(* CODESYS project Example12_PLC.project

Project tree, tasks and I/O mapping:
  Device : CODESYS Control Win V3, 3S - Smart Software Solutions GmbH, order no. 305021, version 3.5.7.0
    application Application
      libraries: Standard, * (System)
      task MainTask (cyclic, interval t#20ms, priority 1) calls PLC_PRG
      program PLC_PRG [ST]
      global variables GVL
      function block FB_G4LTL [ST]
    Ethernet : Ethernet, 3S - Smart Software Solutions GmbH, version 3.5.7.0
      Modbus_TCP_Master : Modbus TCP Master, 3S - Smart Software Solutions GmbH, version 3.5.6.0
          settings: AutoReconnect = TRUE
        Modbus_TCP_Slave : Modbus TCP Slave, 3S - Smart Software Solutions GmbH, version 3.5.7.0
            settings: Unit-ID = 1; IPAddress = [127, 0, 0, 1]; Channel 0.Function Code = 4; Channel 0.Read Offset = 16#0000; Channel 0.Read Length = 1; Channel 0.Write Offset = 0; Channel 0.Write Length = 0; Channel 0.Cycle Time = 100; Channel 1.Function Code = 4; Channel 1.Read Offset = 16#0001; Channel 1.Read Length = 1; Channel 1.Write Offset = 0; Channel 1.Write Length = 0; Channel 1.Cycle Time = 100; Channel 2.Function Code = 4; Channel 2.Read Offset = 16#0002; Channel 2.Read Length = 1; Channel 2.Write Offset = 0; Channel 2.Write Length = 0; Channel 2.Cycle Time = 100; Channel 3.Function Code = 4; Channel 3.Read Offset = 16#0003; Channel 3.Read Length = 1; Channel 3.Write Offset = 0; Channel 3.Write Length = 0; Channel 3.Cycle Time = 100; Channel 4.Function Code = 4; Channel 4.Read Offset = 16#0004; Channel 4.Read Length = 1; Channel 4.Write Offset = 0; Channel 4.Write Length = 0; Channel 4.Cycle Time = 100; Channel 5.Function Code = 6; Channel 5.Read Offset = 0; Channel 5.Read Length = 0; Channel 5.Write Offset = 16#0000; Channel 5.Write Length = 1; Channel 5.Cycle Time = 100; Channel 6.Function Code = 6; Channel 6.Read Offset = 0;
              Channel 6.Read Length = 0; Channel 6.Write Offset = 16#0002; Channel 6.Write Length = 1; Channel 6.Cycle Time = 100; Channel 7.Function Code = 6; Channel 7.Read Offset = 0; Channel 7.Read Length = 0; Channel 7.Write Offset = 16#0003; Channel 7.Write Length = 1; Channel 7.Cycle Time = 100; Channel 8.Function Code = 6; Channel 8.Read Offset = 0; Channel 8.Read Length = 0; Channel 8.Write Offset = 16#0004; Channel 8.Write Length = 1; Channel 8.Cycle Time = 100; Channel 9.Function Code = 6; Channel 9.Read Offset = 0; Channel 9.Read Length = 0; Channel 9.Write Offset = 16#0001; Channel 9.Write Length = 1; Channel 9.Cycle Time = 100; Channel 10.Function Code = 4; Channel 10.Read Offset = 16#0005; Channel 10.Read Length = 1; Channel 10.Write Offset = 0; Channel 10.Write Length = 0; Channel 10.Cycle Time = 100
            input  Application.dIn0 : BOOL  // Channel 0.Channel 0.Bit0
            input  Application.dIn1 : BOOL  // Channel 1.Channel 1.Bit0
            input  Application.dIn2 : BOOL  // Channel 2.Channel 2.Bit0
            input  Application.dIn3 : BOOL  // Channel 3.Channel 3.Bit0
            input  Application.dIn4 : BOOL  // Channel 4.Channel 4.Bit0
            output Application.dOut0 : BOOL  // Channel 5.Channel 5.Bit0
            output Application.dOut2 : BOOL  // Channel 6.Channel 6.Bit0
            output Application.dOut3 : BOOL  // Channel 7.Channel 7.Bit0
            output Application.dOut4 : BOOL  // Channel 8.Channel 8.Bit0
            output Application.dOut1 : BOOL  // Channel 9.Channel 9.Bit0
            input  Application.dIn5 : BOOL  // Channel 10.Channel 10.Bit0
            unmapped channels: Channel 0, Channel 1, Channel 2, Channel 3, Channel 4, Channel 5, Channel 6, Channel 7, Channel 8, Channel 9, Channel 10
*)

// Device/Application/GVL
VAR_GLOBAL
	
dIn0 : BOOL;
dIn1 : BOOL;
dIn2 : BOOL;
dIn3 : BOOL;
dIn4 : BOOL;
dIn5 : BOOL;

dOut0 : BOOL;
dOut1 : BOOL; 
dOut2 : BOOL; 
dOut3 : BOOL; 
dOut4 : BOOL; 
END_VAR

// Device/Application/PLC_PRG
PROGRAM PLC_PRG
 

VAR 
	fb: FB_G4LTL;

	
END_VAR



// Direct looping
// Assign pins (from global variable to function block) 
fb.x0 := dIn0;
fb.x1 := dIn1;
fb.x2 := dIn2;
fb.x3 := dIn3;
fb.x4 := dIn4;
fb.x5 := dIn5;

// Assign pins (from function block to global variable)
dOut0 := fb.y0;
dOut1 := fb.y1;
dOut2 := fb.y2;

// Run the function block
fb();

END_PROGRAM

// Device/Application/FB_G4LTL
FUNCTION_BLOCK FB_G4LTL
   (* Variable definition *)
   VAR_INPUT
      x0	: BOOL;
      x1	: BOOL;
      x2	: BOOL;
      x3	: BOOL;
      x4	: BOOL;
      x5	: BOOL;
   END_VAR
   VAR_OUTPUT
      y0	: BOOL;
      y1	: BOOL;
      y2	: BOOL;
   END_VAR
   VAR
   (* The total number of states equals to 84 *)
      cstate98	: LINT := 0;
   END_VAR
   (* Constant definition  *)

 
   (* Control logic *)
CASE cstate98 OF
2090:
    IF ((x0 = FALSE) AND  (x1 = FALSE) AND  (x2 = FALSE) AND  (x3 = FALSE) AND  ( TRUE ) AND  (x5 = FALSE)) OR ((x0 = FALSE) AND  (x1 = FALSE) AND  (x2 = FALSE) AND  (x3 = TRUE) AND  (x4 = FALSE) AND  (x5 = FALSE)) THEN 
        cstate98 := 2122; y0 := FALSE; y1 := FALSE; y2 := FALSE;  
    ELSIF ((x0 = FALSE) AND  (x1 = FALSE) AND  (x2 = FALSE) AND  (x3 = FALSE) AND  ( TRUE ) AND  (x5 = TRUE)) OR ((x0 = FALSE) AND  (x1 = FALSE) AND  (x2 = FALSE) AND  (x3 = TRUE) AND  (x4 = FALSE) AND  (x5 = TRUE)) THEN 
        cstate98 := 2123; y0 := FALSE; y1 := FALSE; y2 := FALSE;  
    ELSIF ((x0 = FALSE) AND  (x1 = FALSE) AND  (x2 = FALSE) AND  (x3 = TRUE) AND  (x4 = TRUE) AND  ( TRUE )) THEN 
        cstate98 := 2090; y0 := FALSE; y1 := FALSE; y2 := FALSE;  
    ELSIF ((x0 = FALSE) AND  (x1 = FALSE) AND  (x2 = TRUE) AND  (x3 = FALSE) AND  ( TRUE ) AND  (x5 = FALSE)) THEN 
        cstate98 := 2602; y0 := FALSE; y1 := TRUE; y2 := FALSE;  
    ELSIF ((x0 = FALSE) AND  (x1 = FALSE) AND  (x2 = TRUE) AND  (x3 = FALSE) AND  ( TRUE ) AND  (x5 = TRUE)) THEN 
        cstate98 := 1610; y0 := FALSE; y1 := FALSE; y2 := FALSE;  
    ELSIF ((x0 = FALSE) AND  (x1 = FALSE) AND  (x2 = TRUE) AND  (x3 = TRUE) AND  ( TRUE ) AND  ( TRUE )) OR ((x0 = FALSE) AND  (x1 = TRUE) AND  (x2 = FALSE) AND  (x3 = TRUE) AND  ( TRUE ) AND  ( TRUE )) OR ((x0 = FALSE) AND  (x1 = TRUE) AND  (x2 = TRUE) AND  ( TRUE ) AND  ( TRUE ) AND  ( TRUE )) OR ((x0 = TRUE) AND  ( TRUE ) AND  (x2 = FALSE) AND  (x3 = TRUE) AND  ( TRUE ) AND  ( TRUE )) OR ((x0 = TRUE) AND  ( TRUE ) AND  (x2 = TRUE) AND  ( TRUE ) AND  ( TRUE ) AND  ( TRUE )) THEN 
        cstate98 := 617; y0 := FALSE; y1 := FALSE; y2 := FALSE;  
    ELSIF ((x0 = FALSE) AND  (x1 = TRUE) AND  (x2 = FALSE) AND  (x3 = FALSE) AND  ( TRUE ) AND  (x5 = FALSE)) OR ((x0 = TRUE) AND  ( TRUE ) AND  (x2 = FALSE) AND  (x3 = FALSE) AND  ( TRUE ) AND  (x5 = FALSE)) THEN 
        cstate98 := 3210; y0 := TRUE; y1 := FALSE; y2 := FALSE;  
    ELSIF ((x0 = FALSE) AND  (x1 = TRUE) AND  (x2 = FALSE) AND  (x3 = FALSE) AND  ( TRUE ) AND  (x5 = TRUE)) OR ((x0 = TRUE) AND  ( TRUE ) AND  (x2 = FALSE) AND  (x3 = FALSE) AND  ( TRUE ) AND  (x5 = TRUE)) THEN 
        cstate98 := 1194; y0 := FALSE; y1 := FALSE; y2 := FALSE;  
    END_IF;
2608:
    IF ((x0 = FALSE) AND  (x1 = FALSE) AND  (x2 = FALSE) AND  (x3 = FALSE) AND  ( TRUE ) AND  (x5 = FALSE)) OR ((x0 = FALSE) AND  (x1 = FALSE) AND  (x2 = FALSE) AND  (x3 = TRUE) AND  (x4 = FALSE) AND  (x5 = FALSE)) THEN 
        cstate98 := 3632; y0 := FALSE; y1 := TRUE; y2 := FALSE;  
    ELSIF ((x0 = FALSE) AND  (x1 = FALSE) AND  (x2 = FALSE) AND  (x3 = FALSE) AND  ( TRUE ) AND  (x5 = TRUE)) OR ((x0 = FALSE) AND  (x1 = FALSE) AND  (x2 = FALSE) AND  (x3 = TRUE) AND  (x4 = FALSE) AND  (x5 = TRUE)) THEN 
        cstate98 := 2131; y0 := FALSE; y1 := FALSE; y2 := FALSE;  
    ELSIF ((x0 = FALSE) AND  (x1 = FALSE) AND  (x2 = FALSE) AND  (x3 = TRUE) AND  (x4 = TRUE) AND  (x5 = FALSE)) THEN 
        cstate98 := 3624; y0 := FALSE; y1 := TRUE; y2 := FALSE;  
    ELSIF ((x0 = FALSE) AND  (x1 = FALSE) AND  (x2 = FALSE) AND  (x3 = TRUE) AND  (x4 = TRUE) AND  (x5 = TRUE)) THEN 
        cstate98 := 2090; y0 := FALSE; y1 := FALSE; y2 := FALSE;  
    ELSIF ((x0 = FALSE) AND  (x1 = FALSE) AND  (x2 = TRUE) AND  (x3 = FALSE) AND  ( TRUE ) AND  (x5 = FALSE)) THEN 
        cstate98 := 2608; y0 := FALSE; y1 := TRUE; y2 := FALSE;  
    ELSIF ((x0 = FALSE) AND  (x1 = FALSE) AND  (x2 = TRUE) AND  (x3 = FALSE) AND  ( TRUE ) AND  (x5 = TRUE)) THEN 
        cstate98 := 1618; y0 := FALSE; y1 := FALSE; y2 := FALSE;  
    ELSIF ((x0 = FALSE) AND  (x1 = FALSE) AND  (x2 = TRUE) AND  (x3 = TRUE) AND  ( TRUE ) AND  ( TRUE )) OR ((x0 = FALSE) AND  (x1 = TRUE) AND  (x2 = FALSE) AND  (x3 = TRUE) AND  ( TRUE ) AND  ( TRUE )) OR ((x0 = FALSE) AND  (x1 = TRUE) AND  (x2 = TRUE) AND  ( TRUE ) AND  ( TRUE ) AND  ( TRUE )) OR ((x0 = TRUE) AND  ( TRUE ) AND  (x2 = FALSE) AND  (x3 = TRUE) AND  ( TRUE ) AND  ( TRUE )) OR ((x0 = TRUE) AND  ( TRUE ) AND  (x2 = TRUE) AND  ( TRUE ) AND  ( TRUE ) AND  ( TRUE )) THEN 
        cstate98 := 617; y0 := FALSE; y1 := FALSE; y2 := FALSE;  
    ELSIF ((x0 = FALSE) AND  (x1 = TRUE) AND  (x2 = FALSE) AND  (x3 = FALSE) AND  ( TRUE ) AND  (x5 = FALSE)) OR ((x0 = TRUE) AND  ( TRUE ) AND  (x2 = FALSE) AND  (x3 = FALSE) AND  ( TRUE ) AND  (x5 = FALSE)) THEN 
        cstate98 := 3728; y0 := FALSE; y1 := TRUE; y2 := FALSE;  
    ELSIF ((x0 = FALSE) AND  (x1 = TRUE) AND  (x2 = FALSE) AND  (x3 = FALSE) AND  ( TRUE ) AND  (x5 = TRUE)) OR ((x0 = TRUE) AND  ( TRUE ) AND  (x2 = FALSE) AND  (x3 = FALSE) AND  ( TRUE ) AND  (x5 = TRUE)) THEN 
        cstate98 := 1202; y0 := FALSE; y1 := FALSE; y2 := FALSE;  
    END_IF;
2092:
    IF ((x0 = FALSE) AND  (x1 = FALSE) AND  (x2 = FALSE) AND  (x3 = FALSE) AND  ( TRUE ) AND  (x5 = FALSE)) OR ((x0 = FALSE) AND  (x1 = FALSE) AND  (x2 = FALSE) AND  (x3 = TRUE) AND  (x4 = FALSE) AND  (x5 = FALSE)) THEN 
        cstate98 := 2124; y0 := FALSE; y1 := FALSE; y2 := FALSE;  
    ELSIF ((x0 = FALSE) AND  (x1 = FALSE) AND  (x2 = FALSE) AND  (x3 = FALSE) AND  ( TRUE ) AND  (x5 = TRUE)) OR ((x0 = FALSE) AND  (x1 = FALSE) AND  (x2 = FALSE) AND  (x3 = TRUE) AND  (x4 = FALSE) AND  (x5 = TRUE)) THEN 
        cstate98 := 2127; y0 := FALSE; y1 := FALSE; y2 := FALSE;  
    ELSIF ((x0 = FALSE) AND  (x1 = FALSE) AND  (x2 = FALSE) AND  (x3 = TRUE) AND  (x4 = TRUE) AND  (x5 = FALSE)) THEN 
        cstate98 := 2092; y0 := FALSE; y1 := FALSE; y2 := FALSE;  
    ELSIF ((x0 = FALSE) AND  (x1 = FALSE) AND  (x2 = FALSE) AND  (x3 = TRUE) AND  (x4 = TRUE) AND  (x5 = TRUE)) THEN 
        cstate98 := 2094; y0 := FALSE; y1 := FALSE; y2 := FALSE;  
    ELSIF ((x0 = FALSE) AND  (x1 = FALSE) AND  (x2 = TRUE) AND  (x3 = FALSE) AND  ( TRUE ) AND  (x5 = FALSE)) THEN 
        cstate98 := 2600; y0 := FALSE; y1 := TRUE; y2 := FALSE;  
    ELSIF ((x0 = FALSE) AND  (x1 = FALSE) AND  (x2 = TRUE) AND  (x3 = FALSE) AND  ( TRUE ) AND  (x5 = TRUE)) THEN 
        cstate98 := 1610; y0 := FALSE; y1 := FALSE; y2 := FALSE;  
    ELSIF ((x0 = FALSE) AND  (x1 = FALSE) AND  (x2 = TRUE) AND  (x3 = TRUE) AND  ( TRUE ) AND  ( TRUE )) OR ((x0 = FALSE) AND  (x1 = TRUE) AND  (x2 = FALSE) AND  (x3 = TRUE) AND  ( TRUE ) AND  ( TRUE )) OR ((x0 = FALSE) AND  (x1 = TRUE) AND  (x2 = TRUE) AND  ( TRUE ) AND  ( TRUE ) AND  ( TRUE )) OR ((x0 = TRUE) AND  ( TRUE ) AND  (x2 = FALSE) AND  (x3 = TRUE) AND  ( TRUE ) AND  ( TRUE )) OR ((x0 = TRUE) AND  ( TRUE ) AND  (x2 = TRUE) AND  ( TRUE ) AND  ( TRUE ) AND  ( TRUE )) THEN 
        cstate98 := 617; y0 := FALSE; y1 := FALSE; y2 := FALSE;  
    ELSIF ((x0 = FALSE) AND  (x1 = TRUE) AND  (x2 = FALSE) AND  (x3 = FALSE) AND  ( TRUE ) AND  (x5 = FALSE)) OR ((x0 = TRUE) AND  ( TRUE ) AND  (x2 = FALSE) AND  (x3 = FALSE) AND  ( TRUE ) AND  (x5 = FALSE)) THEN 
        cstate98 := 3212; y0 := TRUE; y1 := FALSE; y2 := FALSE;  
    ELSIF ((x0 = FALSE) AND  (x1 = TRUE) AND  (x2 = FALSE) AND  (x3 = FALSE) AND  ( TRUE ) AND  (x5 = TRUE)) OR ((x0 = TRUE) AND  ( TRUE ) AND  (x2 = FALSE) AND  (x3 = FALSE) AND  ( TRUE ) AND  (x5 = TRUE)) THEN 
        cstate98 := 1198; y0 := FALSE; y1 := FALSE; y2 := FALSE;  
    END_IF;
1198:
    IF ((x0 = FALSE) AND  (x1 = FALSE) AND  (x2 = FALSE) AND  (x3 = FALSE) AND  ( TRUE ) AND  (x5 = FALSE)) OR ((x0 = FALSE) AND  (x1 = FALSE) AND  (x2 = FALSE) AND  (x3 = TRUE) AND  (x4 = FALSE) AND  (x5 = FALSE)) THEN 
        cstate98 := 2222; y0 := FALSE; y1 := FALSE; y2 := FALSE;  
    ELSIF ((x0 = FALSE) AND  (x1 = FALSE) AND  (x2 = FALSE) AND  (x3 = FALSE) AND  ( TRUE ) AND  (x5 = TRUE)) OR ((x0 = FALSE) AND  (x1 = FALSE) AND  (x2 = FALSE) AND  (x3 = TRUE) AND  (x4 = FALSE) AND  (x5 = TRUE)) THEN 
        cstate98 := 2223; y0 := FALSE; y1 := FALSE; y2 := FALSE;  
    ELSIF ((x0 = FALSE) AND  (x1 = FALSE) AND  (x2 = FALSE) AND  (x3 = TRUE) AND  (x4 = TRUE) AND  (x5 = FALSE)) THEN 
        cstate98 := 238; y0 := FALSE; y1 := FALSE; y2 := TRUE;  
    ELSIF ((x0 = FALSE) AND  (x1 = FALSE) AND  (x2 = FALSE) AND  (x3 = TRUE) AND  (x4 = TRUE) AND  (x5 = TRUE)) THEN 
        cstate98 := 2190; y0 := FALSE; y1 := FALSE; y2 := FALSE;  
    ELSIF ((x0 = FALSE) AND  (x1 = FALSE) AND  (x2 = TRUE) AND  (x3 = FALSE) AND  ( TRUE ) AND  (x5 = FALSE)) THEN 
        cstate98 := 2698; y0 := FALSE; y1 := TRUE; y2 := FALSE;  
    ELSIF ((x0 = FALSE) AND  (x1 = FALSE) AND  (x2 = TRUE) AND  (x3 = FALSE) AND  ( TRUE ) AND  (x5 = TRUE)) THEN 
        cstate98 := 1706; y0 := FALSE; y1 := FALSE; y2 := FALSE;  
    ELSIF ((x0 = FALSE) AND  (x1 = FALSE) AND  (x2 = TRUE) AND  (x3 = TRUE) AND  ( TRUE ) AND  ( TRUE )) OR ((x0 = FALSE) AND  (x1 = TRUE) AND  (x2 = FALSE) AND  (x3 = TRUE) AND  ( TRUE ) AND  ( TRUE )) OR ((x0 = FALSE) AND  (x1 = TRUE) AND  (x2 = TRUE) AND  ( TRUE ) AND  ( TRUE ) AND  ( TRUE )) OR ((x0 = TRUE) AND  ( TRUE ) AND  (x2 = FALSE) AND  (x3 = TRUE) AND  ( TRUE ) AND  ( TRUE )) OR ((x0 = TRUE) AND  ( TRUE ) AND  (x2 = TRUE) AND  ( TRUE ) AND  ( TRUE ) AND  ( TRUE )) THEN 
        cstate98 := 617; y0 := FALSE; y1 := FALSE; y2 := FALSE;  
    ELSIF ((x0 = FALSE) AND  (x1 = TRUE) AND  (x2 = FALSE) AND  (x3 = FALSE) AND  ( TRUE ) AND  ( TRUE )) OR ((x0 = TRUE) AND  ( TRUE ) AND  (x2 = FALSE) AND  (x3 = FALSE) AND  ( TRUE ) AND  ( TRUE )) THEN 
        cstate98 := 1198; y0 := FALSE; y1 := FALSE; y2 := FALSE;  
    END_IF;
3722:
    IF ((x0 = FALSE) AND  (x1 = FALSE) AND  (x2 = FALSE) AND  ( TRUE ) AND  ( TRUE ) AND  (x5 = FALSE)) OR ((x0 = FALSE) AND  (x1 = TRUE) AND  (x2 = FALSE) AND  (x3 = FALSE) AND  ( TRUE ) AND  (x5 = FALSE)) OR ((x0 = TRUE) AND  ( TRUE ) AND  (x2 = FALSE) AND  (x3 = FALSE) AND  ( TRUE ) AND  (x5 = FALSE)) THEN 
        cstate98 := 3722; y0 := FALSE; y1 := TRUE; y2 := FALSE;  
    ELSIF ((x0 = FALSE) AND  (x1 = FALSE) AND  (x2 = FALSE) AND  (x3 = FALSE) AND  ( TRUE ) AND  (x5 = TRUE)) OR ((x0 = FALSE) AND  (x1 = FALSE) AND  (x2 = FALSE) AND  (x3 = TRUE) AND  (x4 = FALSE) AND  (x5 = TRUE)) THEN 
        cstate98 := 2219; y0 := FALSE; y1 := FALSE; y2 := FALSE;  
    ELSIF ((x0 = FALSE) AND  (x1 = FALSE) AND  (x2 = FALSE) AND  (x3 = TRUE) AND  (x4 = TRUE) AND  (x5 = TRUE)) THEN 
        cstate98 := 2186; y0 := FALSE; y1 := FALSE; y2 := FALSE;  
    ELSIF ((x0 = FALSE) AND  (x1 = FALSE) AND  (x2 = TRUE) AND  (x3 = FALSE) AND  ( TRUE ) AND  (x5 = FALSE)) THEN 
        cstate98 := 2698; y0 := FALSE; y1 := TRUE; y2 := FALSE;  
    ELSIF ((x0 = FALSE) AND  (x1 = FALSE) AND  (x2 = TRUE) AND  (x3 = FALSE) AND  ( TRUE ) AND  (x5 = TRUE)) THEN 
        cstate98 := 1706; y0 := FALSE; y1 := FALSE; y2 := FALSE;  
    ELSIF ((x0 = FALSE) AND  (x1 = FALSE) AND  (x2 = TRUE) AND  (x3 = TRUE) AND  ( TRUE ) AND  ( TRUE )) OR ((x0 = FALSE) AND  (x1 = TRUE) AND  (x2 = FALSE) AND  (x3 = TRUE) AND  ( TRUE ) AND  ( TRUE )) OR ((x0 = FALSE) AND  (x1 = TRUE) AND  (x2 = TRUE) AND  ( TRUE ) AND  ( TRUE ) AND  ( TRUE )) OR ((x0 = TRUE) AND  ( TRUE ) AND  (x2 = FALSE) AND  (x3 = TRUE) AND  ( TRUE ) AND  ( TRUE )) OR ((x0 = TRUE) AND  ( TRUE ) AND  (x2 = TRUE) AND  ( TRUE ) AND  ( TRUE ) AND  ( TRUE )) THEN 
        cstate98 := 617; y0 := FALSE; y1 := FALSE; y2 := FALSE;  
    ELSIF ((x0 = FALSE) AND  (x1 = TRUE) AND  (x2 = FALSE) AND  (x3 = FALSE) AND  ( TRUE ) AND  (x5 = TRUE)) OR ((x0 = TRUE) AND  ( TRUE ) AND  (x2 = FALSE) AND  (x3 = FALSE) AND  ( TRUE ) AND  (x5 = TRUE)) THEN 
        cstate98 := 1194; y0 := FALSE; y1 := FALSE; y2 := FALSE;  
    END_IF;
3720:
    IF ((x0 = FALSE) AND  (x1 = FALSE) AND  (x2 = FALSE) AND  ( TRUE ) AND  ( TRUE ) AND  (x5 = FALSE)) OR ((x0 = FALSE) AND  (x1 = TRUE) AND  (x2 = FALSE) AND  (x3 = FALSE) AND  ( TRUE ) AND  (x5 = FALSE)) OR ((x0 = TRUE) AND  ( TRUE ) AND  (x2 = FALSE) AND  (x3 = FALSE) AND  ( TRUE ) AND  (x5 = FALSE)) THEN 
        cstate98 := 3720; y0 := FALSE; y1 := TRUE; y2 := FALSE;  
    ELSIF ((x0 = FALSE) AND  (x1 = FALSE) AND  (x2 = FALSE) AND  (x3 = FALSE) AND  ( TRUE ) AND  (x5 = TRUE)) OR ((x0 = FALSE) AND  (x1 = FALSE) AND  (x2 = FALSE) AND  (x3 = TRUE) AND  (x4 = FALSE) AND  (x5 = TRUE)) THEN 
        cstate98 := 2219; y0 := FALSE; y1 := FALSE; y2 := FALSE;  
    ELSIF ((x0 = FALSE) AND  (x1 = FALSE) AND  (x2 = FALSE) AND  (x3 = TRUE) AND  (x4 = TRUE) AND  (x5 = TRUE)) THEN 
        cstate98 := 2186; y0 := FALSE; y1 := FALSE; y2 := FALSE;  
    ELSIF ((x0 = FALSE) AND  (x1 = FALSE) AND  (x2 = TRUE) AND  (x3 = FALSE) AND  ( TRUE ) AND  (x5 = FALSE)) THEN 
        cstate98 := 2696; y0 := FALSE; y1 := TRUE; y2 := FALSE;  
    ELSIF ((x0 = FALSE) AND  (x1 = FALSE) AND  (x2 = TRUE) AND  (x3 = FALSE) AND  ( TRUE ) AND  (x5 = TRUE)) THEN 
        cstate98 := 1706; y0 := FALSE; y1 := FALSE; y2 := FALSE;  
    ELSIF ((x0 = FALSE) AND  (x1 = FALSE) AND  (x2 = TRUE) AND  (x3 = TRUE) AND  ( TRUE ) AND  ( TRUE )) OR ((x0 = FALSE) AND  (x1 = TRUE) AND  (x2 = FALSE) AND  (x3 = TRUE) AND  ( TRUE ) AND  ( TRUE )) OR ((x0 = FALSE) AND  (x1 = TRUE) AND  (x2 = TRUE) AND  ( TRUE ) AND  ( TRUE ) AND  ( TRUE )) OR ((x0 = TRUE) AND  ( TRUE ) AND  (x2 = FALSE) AND  (x3 = TRUE) AND  ( TRUE ) AND  ( TRUE )) OR ((x0 = TRUE) AND  ( TRUE ) AND  (x2 = TRUE) AND  ( TRUE ) AND  ( TRUE ) AND  ( TRUE )) THEN 
        cstate98 := 617; y0 := FALSE; y1 := FALSE; y2 := FALSE;  
    ELSIF ((x0 = FALSE) AND  (x1 = TRUE) AND  (x2 = FALSE) AND  (x3 = FALSE) AND  ( TRUE ) AND  (x5 = TRUE)) OR ((x0 = TRUE) AND  ( TRUE ) AND  (x2 = FALSE) AND  (x3 = FALSE) AND  ( TRUE ) AND  (x5 = TRUE)) THEN 
        cstate98 := 1194; y0 := FALSE; y1 := FALSE; y2 := FALSE;  
    END_IF;
1194:
    IF ((x0 = FALSE) AND  (x1 = FALSE) AND  (x2 = FALSE) AND  (x3 = FALSE) AND  ( TRUE ) AND  (x5 = FALSE)) OR ((x0 = FALSE) AND  (x1 = FALSE) AND  (x2 = FALSE) AND  (x3 = TRUE) AND  (x4 = FALSE) AND  (x5 = FALSE)) THEN 
        cstate98 := 2218; y0 := FALSE; y1 := FALSE; y2 := FALSE;  
    ELSIF ((x0 = FALSE) AND  (x1 = FALSE) AND  (x2 = FALSE) AND  (x3 = FALSE) AND  ( TRUE ) AND  (x5 = TRUE)) OR ((x0 = FALSE) AND  (x1 = FALSE) AND  (x2 = FALSE) AND  (x3 = TRUE) AND  (x4 = FALSE) AND  (x5 = TRUE)) THEN 
        cstate98 := 2219; y0 := FALSE; y1 := FALSE; y2 := FALSE;  
    ELSIF ((x0 = FALSE) AND  (x1 = FALSE) AND  (x2 = FALSE) AND  (x3 = TRUE) AND  (x4 = TRUE) AND  (x5 = FALSE)) THEN 
        cstate98 := 234; y0 := FALSE; y1 := FALSE; y2 := TRUE;  
    ELSIF ((x0 = FALSE) AND  (x1 = FALSE) AND  (x2 = FALSE) AND  (x3 = TRUE) AND  (x4 = TRUE) AND  (x5 = TRUE)) THEN 
        cstate98 := 2186; y0 := FALSE; y1 := FALSE; y2 := FALSE;  
    ELSIF ((x0 = FALSE) AND  (x1 = FALSE) AND  (x2 = TRUE) AND  (x3 = FALSE) AND  ( TRUE ) AND  (x5 = FALSE)) THEN 
        cstate98 := 2698; y0 := FALSE; y1 := TRUE; y2 := FALSE;  
    ELSIF ((x0 = FALSE) AND  (x1 = FALSE) AND  (x2 = TRUE) AND  (x3 = FALSE) AND  ( TRUE ) AND  (x5 = TRUE)) THEN 
        cstate98 := 1706; y0 := FALSE; y1 := FALSE; y2 := FALSE;  
    ELSIF ((x0 = FALSE) AND  (x1 = FALSE) AND  (x2 = TRUE) AND  (x3 = TRUE) AND  ( TRUE ) AND  ( TRUE )) OR ((x0 = FALSE) AND  (x1 = TRUE) AND  (x2 = FALSE) AND  (x3 = TRUE) AND  ( TRUE ) AND  ( TRUE )) OR ((x0 = FALSE) AND  (x1 = TRUE) AND  (x2 = TRUE) AND  ( TRUE ) AND  ( TRUE ) AND  ( TRUE )) OR ((x0 = TRUE) AND  ( TRUE ) AND  (x2 = FALSE) AND  (x3 = TRUE) AND  ( TRUE ) AND  ( TRUE )) OR ((x0 = TRUE) AND  ( TRUE ) AND  (x2 = TRUE) AND  ( TRUE ) AND  ( TRUE ) AND  ( TRUE )) THEN 
        cstate98 := 617; y0 := FALSE; y1 := FALSE; y2 := FALSE;  
    ELSIF ((x0 = FALSE) AND  (x1 = TRUE) AND  (x2 = FALSE) AND  (x3 = FALSE) AND  ( TRUE ) AND  ( TRUE )) OR ((x0 = TRUE) AND  ( TRUE ) AND  (x2 = FALSE) AND  (x3 = FALSE) AND  ( TRUE ) AND  ( TRUE )) THEN 
        cstate98 := 1194; y0 := FALSE; y1 := FALSE; y2 := FALSE;  
    END_IF;
2602:
    IF ((x0 = FALSE) AND  (x1 = FALSE) AND  (x2 = FALSE) AND  ( TRUE ) AND  ( TRUE ) AND  (x5 = FALSE)) THEN 
        cstate98 := 3626; y0 := FALSE; y1 := TRUE; y2 := FALSE;  
    ELSIF ((x0 = FALSE) AND  (x1 = FALSE) AND  (x2 = FALSE) AND  (x3 = FALSE) AND  ( TRUE ) AND  (x5 = TRUE)) OR ((x0 = FALSE) AND  (x1 = FALSE) AND  (x2 = FALSE) AND  (x3 = TRUE) AND  (x4 = FALSE) AND  (x5 = TRUE)) THEN 
        cstate98 := 2123; y0 := FALSE; y1 := FALSE; y2 := FALSE;  
    ELSIF ((x0 = FALSE) AND  (x1 = FALSE) AND  (x2 = FALSE) AND  (x3 = TRUE) AND  (x4 = TRUE) AND  (x5 = TRUE)) THEN 
        cstate98 := 2090; y0 := FALSE; y1 := FALSE; y2 := FALSE;  
    ELSIF ((x0 = FALSE) AND  (x1 = FALSE) AND  (x2 = TRUE) AND  (x3 = FALSE) AND  ( TRUE ) AND  (x5 = FALSE)) THEN 
        cstate98 := 2602; y0 := FALSE; y1 := TRUE; y2 := FALSE;  
    ELSIF ((x0 = FALSE) AND  (x1 = FALSE) AND  (x2 = TRUE) AND  (x3 = FALSE) AND  ( TRUE ) AND  (x5 = TRUE)) THEN 
        cstate98 := 1610; y0 := FALSE; y1 := FALSE; y2 := FALSE;  
    ELSIF ((x0 = FALSE) AND  (x1 = FALSE) AND  (x2 = TRUE) AND  (x3 = TRUE) AND  ( TRUE ) AND  ( TRUE )) OR ((x0 = FALSE) AND  (x1 = TRUE) AND  (x2 = FALSE) AND  (x3 = TRUE) AND  ( TRUE ) AND  ( TRUE )) OR ((x0 = FALSE) AND  (x1 = TRUE) AND  (x2 = TRUE) AND  ( TRUE ) AND  ( TRUE ) AND  ( TRUE )) OR ((x0 = TRUE) AND  ( TRUE ) AND  (x2 = FALSE) AND  (x3 = TRUE) AND  ( TRUE ) AND  ( TRUE )) OR ((x0 = TRUE) AND  ( TRUE ) AND  (x2 = TRUE) AND  ( TRUE ) AND  ( TRUE ) AND  ( TRUE )) THEN 
        cstate98 := 617; y0 := FALSE; y1 := FALSE; y2 := FALSE;  
    ELSIF ((x0 = FALSE) AND  (x1 = TRUE) AND  (x2 = FALSE) AND  (x3 = FALSE) AND  ( TRUE ) AND  (x5 = FALSE)) OR ((x0 = TRUE) AND  ( TRUE ) AND  (x2 = FALSE) AND  (x3 = FALSE) AND  ( TRUE ) AND  (x5 = FALSE)) THEN 
        cstate98 := 3722; y0 := FALSE; y1 := TRUE; y2 := FALSE;  
    ELSIF ((x0 = FALSE) AND  (x1 = TRUE) AND  (x2 = FALSE) AND  (x3 = FALSE) AND  ( TRUE ) AND  (x5 = TRUE)) OR ((x0 = TRUE) AND  ( TRUE ) AND  (x2 = FALSE) AND  (x3 = FALSE) AND  ( TRUE ) AND  (x5 = TRUE)) THEN 
        cstate98 := 1194; y0 := FALSE; y1 := FALSE; y2 := FALSE;  
    END_IF;
2706:
    IF ((x0 = FALSE) AND  (x1 = FALSE) AND  (x2 = FALSE) AND  (x3 = FALSE) AND  ( TRUE ) AND  (x5 = FALSE)) OR ((x0 = FALSE) AND  (x1 = FALSE) AND  (x2 = FALSE) AND  (x3 = TRUE) AND  (x4 = FALSE) AND  (x5 = FALSE)) OR ((x0 = FALSE) AND  (x1 = TRUE) AND  (x2 = FALSE) AND  (x3 = FALSE) AND  ( TRUE ) AND  (x5 = FALSE)) OR ((x0 = TRUE) AND  ( TRUE ) AND  (x2 = FALSE) AND  (x3 = FALSE) AND  ( TRUE ) AND  (x5 = FALSE)) THEN 
        cstate98 := 3730; y0 := FALSE; y1 := TRUE; y2 := FALSE;  
    ELSIF ((x0 = FALSE) AND  (x1 = FALSE) AND  (x2 = FALSE) AND  (x3 = FALSE) AND  ( TRUE ) AND  (x5 = TRUE)) OR ((x0 = FALSE) AND  (x1 = FALSE) AND  (x2 = FALSE) AND  (x3 = TRUE) AND  (x4 = FALSE) AND  (x5 = TRUE)) THEN 
        cstate98 := 2227; y0 := FALSE; y1 := FALSE; y2 := FALSE;  
    ELSIF ((x0 = FALSE) AND  (x1 = FALSE) AND  (x2 = FALSE) AND  (x3 = TRUE) AND  (x4 = TRUE) AND  (x5 = FALSE)) THEN 
        cstate98 := 3722; y0 := FALSE; y1 := TRUE; y2 := FALSE;  
    ELSIF ((x0 = FALSE) AND  (x1 = FALSE) AND  (x2 = FALSE) AND  (x3 = TRUE) AND  (x4 = TRUE) AND  (x5 = TRUE)) THEN 
        cstate98 := 2186; y0 := FALSE; y1 := FALSE; y2 := FALSE;  
    ELSIF ((x0 = FALSE) AND  (x1 = FALSE) AND  (x2 = TRUE) AND  (x3 = FALSE) AND  ( TRUE ) AND  (x5 = FALSE)) THEN 
        cstate98 := 2706; y0 := FALSE; y1 := TRUE; y2 := FALSE;  
    ELSIF ((x0 = FALSE) AND  (x1 = FALSE) AND  (x2 = TRUE) AND  (x3 = FALSE) AND  ( TRUE ) AND  (x5 = TRUE)) THEN 
        cstate98 := 1714; y0 := FALSE; y1 := FALSE; y2 := FALSE;  
    ELSIF ((x0 = FALSE) AND  (x1 = FALSE) AND  (x2 = TRUE) AND  (x3 = TRUE) AND  ( TRUE ) AND  ( TRUE )) OR ((x0 = FALSE) AND  (x1 = TRUE) AND  (x2 = FALSE) AND  (x3 = TRUE) AND  ( TRUE ) AND  ( TRUE )) OR ((x0 = FALSE) AND  (x1 = TRUE) AND  (x2 = TRUE) AND  ( TRUE ) AND  ( TRUE ) AND  ( TRUE )) OR ((x0 = TRUE) AND  ( TRUE ) AND  (x2 = FALSE) AND  (x3 = TRUE) AND  ( TRUE ) AND  ( TRUE )) OR ((x0 = TRUE) AND  ( TRUE ) AND  (x2 = TRUE) AND  ( TRUE ) AND  ( TRUE ) AND  ( TRUE )) THEN 
        cstate98 := 617; y0 := FALSE; y1 := FALSE; y2 := FALSE;  
    ELSIF ((x0 = FALSE) AND  (x1 = TRUE) AND  (x2 = FALSE) AND  (x3 = FALSE) AND  ( TRUE ) AND  (x5 = TRUE)) OR ((x0 = TRUE) AND  ( TRUE ) AND  (x2 = FALSE) AND  (x3 = FALSE) AND  ( TRUE ) AND  (x5 = TRUE)) THEN 
        cstate98 := 1202; y0 := FALSE; y1 := FALSE; y2 := FALSE;  
    END_IF;
2600:
    IF ((x0 = FALSE) AND  (x1 = FALSE) AND  (x2 = FALSE) AND  ( TRUE ) AND  ( TRUE ) AND  (x5 = FALSE)) THEN 
        cstate98 := 3624; y0 := FALSE; y1 := TRUE; y2 := FALSE;  
    ELSIF ((x0 = FALSE) AND  (x1 = FALSE) AND  (x2 = FALSE) AND  (x3 = FALSE) AND  ( TRUE ) AND  (x5 = TRUE)) OR ((x0 = FALSE) AND  (x1 = FALSE) AND  (x2 = FALSE) AND  (x3 = TRUE) AND  (x4 = FALSE) AND  (x5 = TRUE)) THEN 
        cstate98 := 2123; y0 := FALSE; y1 := FALSE; y2 := FALSE;  
    ELSIF ((x0 = FALSE) AND  (x1 = FALSE) AND  (x2 = FALSE) AND  (x3 = TRUE) AND  (x4 = TRUE) AND  (x5 = TRUE)) THEN 
        cstate98 := 2090; y0 := FALSE; y1 := FALSE; y2 := FALSE;  
    ELSIF ((x0 = FALSE) AND  (x1 = FALSE) AND  (x2 = TRUE) AND  (x3 = FALSE) AND  ( TRUE ) AND  (x5 = FALSE)) THEN 
        cstate98 := 2600; y0 := FALSE; y1 := TRUE; y2 := FALSE;  
    ELSIF ((x0 = FALSE) AND  (x1 = FALSE) AND  (x2 = TRUE) AND  (x3 = FALSE) AND  ( TRUE ) AND  (x5 = TRUE)) THEN 
        cstate98 := 1610; y0 := FALSE; y1 := FALSE; y2 := FALSE;  
    ELSIF ((x0 = FALSE) AND  (x1 = FALSE) AND  (x2 = TRUE) AND  (x3 = TRUE) AND  ( TRUE ) AND  ( TRUE )) OR ((x0 = FALSE) AND  (x1 = TRUE) AND  (x2 = FALSE) AND  (x3 = TRUE) AND  ( TRUE ) AND  ( TRUE )) OR ((x0 = FALSE) AND  (x1 = TRUE) AND  (x2 = TRUE) AND  ( TRUE ) AND  ( TRUE ) AND  ( TRUE )) OR ((x0 = TRUE) AND  ( TRUE ) AND  (x2 = FALSE) AND  (x3 = TRUE) AND  ( TRUE ) AND  ( TRUE )) OR ((x0 = TRUE) AND  ( TRUE ) AND  (x2 = TRUE) AND  ( TRUE ) AND  ( TRUE ) AND  ( TRUE )) THEN 
        cstate98 := 617; y0 := FALSE; y1 := FALSE; y2 := FALSE;  
    ELSIF ((x0 = FALSE) AND  (x1 = TRUE) AND  (x2 = FALSE) AND  (x3 = FALSE) AND  ( TRUE ) AND  (x5 = FALSE)) OR ((x0 = TRUE) AND  ( TRUE ) AND  (x2 = FALSE) AND  (x3 = FALSE) AND  ( TRUE ) AND  (x5 = FALSE)) THEN 
        cstate98 := 3720; y0 := FALSE; y1 := TRUE; y2 := FALSE;  
    ELSIF ((x0 = FALSE) AND  (x1 = TRUE) AND  (x2 = FALSE) AND  (x3 = FALSE) AND  ( TRUE ) AND  (x5 = TRUE)) OR ((x0 = TRUE) AND  ( TRUE ) AND  (x2 = FALSE) AND  (x3 = FALSE) AND  ( TRUE ) AND  (x5 = TRUE)) THEN 
        cstate98 := 1194; y0 := FALSE; y1 := FALSE; y2 := FALSE;  
    END_IF;
1190:
    IF ((x0 = FALSE) AND  (x1 = FALSE) AND  (x2 = FALSE) AND  (x3 = FALSE) AND  ( TRUE ) AND  (x5 = FALSE)) OR ((x0 = FALSE) AND  (x1 = FALSE) AND  (x2 = FALSE) AND  (x3 = TRUE) AND  (x4 = FALSE) AND  (x5 = FALSE)) THEN 
        cstate98 := 2214; y0 := FALSE; y1 := FALSE; y2 := FALSE;  
    ELSIF ((x0 = FALSE) AND  (x1 = FALSE) AND  (x2 = FALSE) AND  (x3 = FALSE) AND  ( TRUE ) AND  (x5 = TRUE)) OR ((x0 = FALSE) AND  (x1 = FALSE) AND  (x2 = FALSE) AND  (x3 = TRUE) AND  (x4 = FALSE) AND  (x5 = TRUE)) THEN 
        cstate98 := 2215; y0 := FALSE; y1 := FALSE; y2 := FALSE;  
    ELSIF ((x0 = FALSE) AND  (x1 = FALSE) AND  (x2 = FALSE) AND  (x3 = TRUE) AND  (x4 = TRUE) AND  (x5 = FALSE)) THEN 
        cstate98 := 238; y0 := FALSE; y1 := FALSE; y2 := TRUE;  
    ELSIF ((x0 = FALSE) AND  (x1 = FALSE) AND  (x2 = FALSE) AND  (x3 = TRUE) AND  (x4 = TRUE) AND  (x5 = TRUE)) THEN 
        cstate98 := 2190; y0 := FALSE; y1 := FALSE; y2 := FALSE;  
    ELSIF ((x0 = FALSE) AND  (x1 = FALSE) AND  (x2 = TRUE) AND  (x3 = FALSE) AND  ( TRUE ) AND  (x5 = FALSE)) THEN 
        cstate98 := 2706; y0 := FALSE; y1 := TRUE; y2 := FALSE;  
    ELSIF ((x0 = FALSE) AND  (x1 = FALSE) AND  (x2 = TRUE) AND  (x3 = FALSE) AND  ( TRUE ) AND  (x5 = TRUE)) THEN 
        cstate98 := 1714; y0 := FALSE; y1 := FALSE; y2 := FALSE;  
    ELSIF ((x0 = FALSE) AND  (x1 = FALSE) AND  (x2 = TRUE) AND  (x3 = TRUE) AND  ( TRUE ) AND  ( TRUE )) OR ((x0 = FALSE) AND  (x1 = TRUE) AND  (x2 = FALSE) AND  (x3 = TRUE) AND  ( TRUE ) AND  ( TRUE )) OR ((x0 = FALSE) AND  (x1 = TRUE) AND  (x2 = TRUE) AND  ( TRUE ) AND  ( TRUE ) AND  ( TRUE )) OR ((x0 = TRUE) AND  ( TRUE ) AND  (x2 = FALSE) AND  (x3 = TRUE) AND  ( TRUE ) AND  ( TRUE )) OR ((x0 = TRUE) AND  ( TRUE ) AND  (x2 = TRUE) AND  ( TRUE ) AND  ( TRUE ) AND  ( TRUE )) THEN 
        cstate98 := 617; y0 := FALSE; y1 := FALSE; y2 := FALSE;  
    ELSIF ((x0 = FALSE) AND  (x1 = TRUE) AND  (x2 = FALSE) AND  (x3 = FALSE) AND  ( TRUE ) AND  ( TRUE )) OR ((x0 = TRUE) AND  ( TRUE ) AND  (x2 = FALSE) AND  (x3 = FALSE) AND  ( TRUE ) AND  ( TRUE )) THEN 
        cstate98 := 1190; y0 := FALSE; y1 := FALSE; y2 := FALSE;  
    END_IF;
2704:
    IF ((x0 = FALSE) AND  (x1 = FALSE) AND  (x2 = FALSE) AND  (x3 = FALSE) AND  ( TRUE ) AND  (x5 = FALSE)) OR ((x0 = FALSE) AND  (x1 = FALSE) AND  (x2 = FALSE) AND  (x3 = TRUE) AND  (x4 = FALSE) AND  (x5 = FALSE)) OR ((x0 = FALSE) AND  (x1 = TRUE) AND  (x2 = FALSE) AND  (x3 = FALSE) AND  ( TRUE ) AND  (x5 = FALSE)) OR ((x0 = TRUE) AND  ( TRUE ) AND  (x2 = FALSE) AND  (x3 = FALSE) AND  ( TRUE ) AND  (x5 = FALSE)) THEN 
        cstate98 := 3728; y0 := FALSE; y1 := TRUE; y2 := FALSE;  
    ELSIF ((x0 = FALSE) AND  (x1 = FALSE) AND  (x2 = FALSE) AND  (x3 = FALSE) AND  ( TRUE ) AND  (x5 = TRUE)) OR ((x0 = FALSE) AND  (x1 = FALSE) AND  (x2 = FALSE) AND  (x3 = TRUE) AND  (x4 = FALSE) AND  (x5 = TRUE)) THEN 
        cstate98 := 2227; y0 := FALSE; y1 := FALSE; y2 := FALSE;  
    ELSIF ((x0 = FALSE) AND  (x1 = FALSE) AND  (x2 = FALSE) AND  (x3 = TRUE) AND  (x4 = TRUE) AND  (x5 = FALSE)) THEN 
        cstate98 := 3720; y0 := FALSE; y1 := TRUE; y2 := FALSE;  
    ELSIF ((x0 = FALSE) AND  (x1 = FALSE) AND  (x2 = FALSE) AND  (x3 = TRUE) AND  (x4 = TRUE) AND  (x5 = TRUE)) THEN 
        cstate98 := 2186; y0 := FALSE; y1 := FALSE; y2 := FALSE;  
    ELSIF ((x0 = FALSE) AND  (x1 = FALSE) AND  (x2 = TRUE) AND  (x3 = FALSE) AND  ( TRUE ) AND  (x5 = FALSE)) THEN 
        cstate98 := 2704; y0 := FALSE; y1 := TRUE; y2 := FALSE;  
    ELSIF ((x0 = FALSE) AND  (x1 = FALSE) AND  (x2 = TRUE) AND  (x3 = FALSE) AND  ( TRUE ) AND  (x5 = TRUE)) THEN 
        cstate98 := 1714; y0 := FALSE; y1 := FALSE; y2 := FALSE;  
    ELSIF ((x0 = FALSE) AND  (x1 = FALSE) AND  (x2 = TRUE) AND  (x3 = TRUE) AND  ( TRUE ) AND  ( TRUE )) OR ((x0 = FALSE) AND  (x1 = TRUE) AND  (x2 = FALSE) AND  (x3 = TRUE) AND  ( TRUE ) AND  ( TRUE )) OR ((x0 = FALSE) AND  (x1 = TRUE) AND  (x2 = TRUE) AND  ( TRUE ) AND  ( TRUE ) AND  ( TRUE )) OR ((x0 = TRUE) AND  ( TRUE ) AND  (x2 = FALSE) AND  (x3 = TRUE) AND  ( TRUE ) AND  ( TRUE )) OR ((x0 = TRUE) AND  ( TRUE ) AND  (x2 = TRUE) AND  ( TRUE ) AND  ( TRUE ) AND  ( TRUE )) THEN 
        cstate98 := 617; y0 := FALSE; y1 := FALSE; y2 := FALSE;  
    ELSIF ((x0 = FALSE) AND  (x1 = TRUE) AND  (x2 = FALSE) AND  (x3 = FALSE) AND  ( TRUE ) AND  (x5 = TRUE)) OR ((x0 = TRUE) AND  ( TRUE ) AND  (x2 = FALSE) AND  (x3 = FALSE) AND  ( TRUE ) AND  (x5 = TRUE)) THEN 
        cstate98 := 1202; y0 := FALSE; y1 := FALSE; y2 := FALSE;  
    END_IF;
2094:
    IF ((x0 = FALSE) AND  (x1 = FALSE) AND  (x2 = FALSE) AND  (x3 = FALSE) AND  ( TRUE ) AND  (x5 = FALSE)) OR ((x0 = FALSE) AND  (x1 = FALSE) AND  (x2 = FALSE) AND  (x3 = TRUE) AND  (x4 = FALSE) AND  (x5 = FALSE)) THEN 
        cstate98 := 2126; y0 := FALSE; y1 := FALSE; y2 := FALSE;  
    ELSIF ((x0 = FALSE) AND  (x1 = FALSE) AND  (x2 = FALSE) AND  (x3 = FALSE) AND  ( TRUE ) AND  (x5 = TRUE)) OR ((x0 = FALSE) AND  (x1 = FALSE) AND  (x2 = FALSE) AND  (x3 = TRUE) AND  (x4 = FALSE) AND  (x5 = TRUE)) THEN 
        cstate98 := 2127; y0 := FALSE; y1 := FALSE; y2 := FALSE;  
    ELSIF ((x0 = FALSE) AND  (x1 = FALSE) AND  (x2 = FALSE) AND  (x3 = TRUE) AND  (x4 = TRUE) AND  ( TRUE )) THEN 
        cstate98 := 2094; y0 := FALSE; y1 := FALSE; y2 := FALSE;  
    ELSIF ((x0 = FALSE) AND  (x1 = FALSE) AND  (x2 = TRUE) AND  (x3 = FALSE) AND  ( TRUE ) AND  (x5 = FALSE)) THEN 
        cstate98 := 2602; y0 := FALSE; y1 := TRUE; y2 := FALSE;  
    ELSIF ((x0 = FALSE) AND  (x1 = FALSE) AND  (x2 = TRUE) AND  (x3 = FALSE) AND  ( TRUE ) AND  (x5 = TRUE)) THEN 
        cstate98 := 1610; y0 := FALSE; y1 := FALSE; y2 := FALSE;  
    ELSIF ((x0 = FALSE) AND  (x1 = FALSE) AND  (x2 = TRUE) AND  (x3 = TRUE) AND  ( TRUE ) AND  ( TRUE )) OR ((x0 = FALSE) AND  (x1 = TRUE) AND  (x2 = FALSE) AND  (x3 = TRUE) AND  ( TRUE ) AND  ( TRUE )) OR ((x0 = FALSE) AND  (x1 = TRUE) AND  (x2 = TRUE) AND  ( TRUE ) AND  ( TRUE ) AND  ( TRUE )) OR ((x0 = TRUE) AND  ( TRUE ) AND  (x2 = FALSE) AND  (x3 = TRUE) AND  ( TRUE ) AND  ( TRUE )) OR ((x0 = TRUE) AND  ( TRUE ) AND  (x2 = TRUE) AND  ( TRUE ) AND  ( TRUE ) AND  ( TRUE )) THEN 
        cstate98 := 617; y0 := FALSE; y1 := FALSE; y2 := FALSE;  
    ELSIF ((x0 = FALSE) AND  (x1 = TRUE) AND  (x2 = FALSE) AND  (x3 = FALSE) AND  ( TRUE ) AND  (x5 = FALSE)) OR ((x0 = TRUE) AND  ( TRUE ) AND  (x2 = FALSE) AND  (x3 = FALSE) AND  ( TRUE ) AND  (x5 = FALSE)) THEN 
        cstate98 := 3214; y0 := TRUE; y1 := FALSE; y2 := FALSE;  
    ELSIF ((x0 = FALSE) AND  (x1 = TRUE) AND  (x2 = FALSE) AND  (x3 = FALSE) AND  ( TRUE ) AND  (x5 = TRUE)) OR ((x0 = TRUE) AND  ( TRUE ) AND  (x2 = FALSE) AND  (x3 = FALSE) AND  ( TRUE ) AND  (x5 = TRUE)) THEN 
        cstate98 := 1198; y0 := FALSE; y1 := FALSE; y2 := FALSE;  
    END_IF;
3728:
    IF ((x0 = FALSE) AND  (x1 = FALSE) AND  (x2 = FALSE) AND  (x3 = FALSE) AND  ( TRUE ) AND  (x5 = FALSE)) OR ((x0 = FALSE) AND  (x1 = FALSE) AND  (x2 = FALSE) AND  (x3 = TRUE) AND  (x4 = FALSE) AND  (x5 = FALSE)) OR ((x0 = FALSE) AND  (x1 = TRUE) AND  (x2 = FALSE) AND  (x3 = FALSE) AND  ( TRUE ) AND  (x5 = FALSE)) OR ((x0 = TRUE) AND  ( TRUE ) AND  (x2 = FALSE) AND  (x3 = FALSE) AND  ( TRUE ) AND  (x5 = FALSE)) THEN 
        cstate98 := 3728; y0 := FALSE; y1 := TRUE; y2 := FALSE;  
    ELSIF ((x0 = FALSE) AND  (x1 = FALSE) AND  (x2 = FALSE) AND  (x3 = FALSE) AND  ( TRUE ) AND  (x5 = TRUE)) OR ((x0 = FALSE) AND  (x1 = FALSE) AND  (x2 = FALSE) AND  (x3 = TRUE) AND  (x4 = FALSE) AND  (x5 = TRUE)) THEN 
        cstate98 := 2227; y0 := FALSE; y1 := FALSE; y2 := FALSE;  
    ELSIF ((x0 = FALSE) AND  (x1 = FALSE) AND  (x2 = FALSE) AND  (x3 = TRUE) AND  (x4 = TRUE) AND  (x5 = FALSE)) THEN 
        cstate98 := 3720; y0 := FALSE; y1 := TRUE; y2 := FALSE;  
    ELSIF ((x0 = FALSE) AND  (x1 = FALSE) AND  (x2 = FALSE) AND  (x3 = TRUE) AND  (x4 = TRUE) AND  (x5 = TRUE)) THEN 
        cstate98 := 2186; y0 := FALSE; y1 := FALSE; y2 := FALSE;  
    ELSIF ((x0 = FALSE) AND  (x1 = FALSE) AND  (x2 = TRUE) AND  (x3 = FALSE) AND  ( TRUE ) AND  (x5 = FALSE)) THEN 
        cstate98 := 2704; y0 := FALSE; y1 := TRUE; y2 := FALSE;  
    ELSIF ((x0 = FALSE) AND  (x1 = FALSE) AND  (x2 = TRUE) AND  (x3 = FALSE) AND  ( TRUE ) AND  (x5 = TRUE)) THEN 
        cstate98 := 1714; y0 := FALSE; y1 := FALSE; y2 := FALSE;  
    ELSIF ((x0 = FALSE) AND  (x1 = FALSE) AND  (x2 = TRUE) AND  (x3 = TRUE) AND  ( TRUE ) AND  ( TRUE )) OR ((x0 = FALSE) AND  (x1 = TRUE) AND  (x2 = FALSE) AND  (x3 = TRUE) AND  ( TRUE ) AND  ( TRUE )) OR ((x0 = FALSE) AND  (x1 = TRUE) AND  (x2 = TRUE) AND  ( TRUE ) AND  ( TRUE ) AND  ( TRUE )) OR ((x0 = TRUE) AND  ( TRUE ) AND  (x2 = FALSE) AND  (x3 = TRUE) AND  ( TRUE ) AND  ( TRUE )) OR ((x0 = TRUE) AND  ( TRUE ) AND  (x2 = TRUE) AND  ( TRUE ) AND  ( TRUE ) AND  ( TRUE )) THEN 
        cstate98 := 617; y0 := FALSE; y1 := FALSE; y2 := FALSE;  
    ELSIF ((x0 = FALSE) AND  (x1 = TRUE) AND  (x2 = FALSE) AND  (x3 = FALSE) AND  ( TRUE ) AND  (x5 = TRUE)) OR ((x0 = TRUE) AND  ( TRUE ) AND  (x2 = FALSE) AND  (x3 = FALSE) AND  ( TRUE ) AND  (x5 = TRUE)) THEN 
        cstate98 := 1202; y0 := FALSE; y1 := FALSE; y2 := FALSE;  
    END_IF;
3626:
    IF ((x0 = FALSE) AND  (x1 = FALSE) AND  (x2 = FALSE) AND  ( TRUE ) AND  ( TRUE ) AND  (x5 = FALSE)) THEN 
        cstate98 := 3626; y0 := FALSE; y1 := TRUE; y2 := FALSE;  
    ELSIF ((x0 = FALSE) AND  (x1 = FALSE) AND  (x2 = FALSE) AND  (x3 = FALSE) AND  ( TRUE ) AND  (x5 = TRUE)) OR ((x0 = FALSE) AND  (x1 = FALSE) AND  (x2 = FALSE) AND  (x3 = TRUE) AND  (x4 = FALSE) AND  (x5 = TRUE)) THEN 
        cstate98 := 2123; y0 := FALSE; y1 := FALSE; y2 := FALSE;  
    ELSIF ((x0 = FALSE) AND  (x1 = FALSE) AND  (x2 = FALSE) AND  (x3 = TRUE) AND  (x4 = TRUE) AND  (x5 = TRUE)) THEN 
        cstate98 := 2090; y0 := FALSE; y1 := FALSE; y2 := FALSE;  
    ELSIF ((x0 = FALSE) AND  (x1 = FALSE) AND  (x2 = TRUE) AND  (x3 = FALSE) AND  ( TRUE ) AND  (x5 = FALSE)) THEN 
        cstate98 := 2602; y0 := FALSE; y1 := TRUE; y2 := FALSE;  
    ELSIF ((x0 = FALSE) AND  (x1 = FALSE) AND  (x2 = TRUE) AND  (x3 = FALSE) AND  ( TRUE ) AND  (x5 = TRUE)) THEN 
        cstate98 := 1610; y0 := FALSE; y1 := FALSE; y2 := FALSE;  
    ELSIF ((x0 = FALSE) AND  (x1 = FALSE) AND  (x2 = TRUE) AND  (x3 = TRUE) AND  ( TRUE ) AND  ( TRUE )) OR ((x0 = FALSE) AND  (x1 = TRUE) AND  (x2 = FALSE) AND  (x3 = TRUE) AND  ( TRUE ) AND  ( TRUE )) OR ((x0 = FALSE) AND  (x1 = TRUE) AND  (x2 = TRUE) AND  ( TRUE ) AND  ( TRUE ) AND  ( TRUE )) OR ((x0 = TRUE) AND  ( TRUE ) AND  (x2 = FALSE) AND  (x3 = TRUE) AND  ( TRUE ) AND  ( TRUE )) OR ((x0 = TRUE) AND  ( TRUE ) AND  (x2 = TRUE) AND  ( TRUE ) AND  ( TRUE ) AND  ( TRUE )) THEN 
        cstate98 := 617; y0 := FALSE; y1 := FALSE; y2 := FALSE;  
    ELSIF ((x0 = FALSE) AND  (x1 = TRUE) AND  (x2 = FALSE) AND  (x3 = FALSE) AND  ( TRUE ) AND  (x5 = FALSE)) OR ((x0 = TRUE) AND  ( TRUE ) AND  (x2 = FALSE) AND  (x3 = FALSE) AND  ( TRUE ) AND  (x5 = FALSE)) THEN 
        cstate98 := 3722; y0 := FALSE; y1 := TRUE; y2 := FALSE;  
    ELSIF ((x0 = FALSE) AND  (x1 = TRUE) AND  (x2 = FALSE) AND  (x3 = FALSE) AND  ( TRUE ) AND  (x5 = TRUE)) OR ((x0 = TRUE) AND  ( TRUE ) AND  (x2 = FALSE) AND  (x3 = FALSE) AND  ( TRUE ) AND  (x5 = TRUE)) THEN 
        cstate98 := 1194; y0 := FALSE; y1 := FALSE; y2 := FALSE;  
    END_IF;
3624:
    IF ((x0 = FALSE) AND  (x1 = FALSE) AND  (x2 = FALSE) AND  ( TRUE ) AND  ( TRUE ) AND  (x5 = FALSE)) THEN 
        cstate98 := 3624; y0 := FALSE; y1 := TRUE; y2 := FALSE;  
    ELSIF ((x0 = FALSE) AND  (x1 = FALSE) AND  (x2 = FALSE) AND  (x3 = FALSE) AND  ( TRUE ) AND  (x5 = TRUE)) OR ((x0 = FALSE) AND  (x1 = FALSE) AND  (x2 = FALSE) AND  (x3 = TRUE) AND  (x4 = FALSE) AND  (x5 = TRUE)) THEN 
        cstate98 := 2123; y0 := FALSE; y1 := FALSE; y2 := FALSE;  
    ELSIF ((x0 = FALSE) AND  (x1 = FALSE) AND  (x2 = FALSE) AND  (x3 = TRUE) AND  (x4 = TRUE) AND  (x5 = TRUE)) THEN 
        cstate98 := 2090; y0 := FALSE; y1 := FALSE; y2 := FALSE;  
    ELSIF ((x0 = FALSE) AND  (x1 = FALSE) AND  (x2 = TRUE) AND  (x3 = FALSE) AND  ( TRUE ) AND  (x5 = FALSE)) THEN 
        cstate98 := 2600; y0 := FALSE; y1 := TRUE; y2 := FALSE;  
    ELSIF ((x0 = FALSE) AND  (x1 = FALSE) AND  (x2 = TRUE) AND  (x3 = FALSE) AND  ( TRUE ) AND  (x5 = TRUE)) THEN 
        cstate98 := 1610; y0 := FALSE; y1 := FALSE; y2 := FALSE;  
    ELSIF ((x0 = FALSE) AND  (x1 = FALSE) AND  (x2 = TRUE) AND  (x3 = TRUE) AND  ( TRUE ) AND  ( TRUE )) OR ((x0 = FALSE) AND  (x1 = TRUE) AND  (x2 = FALSE) AND  (x3 = TRUE) AND  ( TRUE ) AND  ( TRUE )) OR ((x0 = FALSE) AND  (x1 = TRUE) AND  (x2 = TRUE) AND  ( TRUE ) AND  ( TRUE ) AND  ( TRUE )) OR ((x0 = TRUE) AND  ( TRUE ) AND  (x2 = FALSE) AND  (x3 = TRUE) AND  ( TRUE ) AND  ( TRUE )) OR ((x0 = TRUE) AND  ( TRUE ) AND  (x2 = TRUE) AND  ( TRUE ) AND  ( TRUE ) AND  ( TRUE )) THEN 
        cstate98 := 617; y0 := FALSE; y1 := FALSE; y2 := FALSE;  
    ELSIF ((x0 = FALSE) AND  (x1 = TRUE) AND  (x2 = FALSE) AND  (x3 = FALSE) AND  ( TRUE ) AND  (x5 = FALSE)) OR ((x0 = TRUE) AND  ( TRUE ) AND  (x2 = FALSE) AND  (x3 = FALSE) AND  ( TRUE ) AND  (x5 = FALSE)) THEN 
        cstate98 := 3720; y0 := FALSE; y1 := TRUE; y2 := FALSE;  
    ELSIF ((x0 = FALSE) AND  (x1 = TRUE) AND  (x2 = FALSE) AND  (x3 = FALSE) AND  ( TRUE ) AND  (x5 = TRUE)) OR ((x0 = TRUE) AND  ( TRUE ) AND  (x2 = FALSE) AND  (x3 = FALSE) AND  ( TRUE ) AND  (x5 = TRUE)) THEN 
        cstate98 := 1194; y0 := FALSE; y1 := FALSE; y2 := FALSE;  
    END_IF;
3632:
    IF ((x0 = FALSE) AND  (x1 = FALSE) AND  (x2 = FALSE) AND  (x3 = FALSE) AND  ( TRUE ) AND  (x5 = FALSE)) OR ((x0 = FALSE) AND  (x1 = FALSE) AND  (x2 = FALSE) AND  (x3 = TRUE) AND  (x4 = FALSE) AND  (x5 = FALSE)) THEN 
        cstate98 := 3632; y0 := FALSE; y1 := TRUE; y2 := FALSE;  
    ELSIF ((x0 = FALSE) AND  (x1 = FALSE) AND  (x2 = FALSE) AND  (x3 = FALSE) AND  ( TRUE ) AND  (x5 = TRUE)) OR ((x0 = FALSE) AND  (x1 = FALSE) AND  (x2 = FALSE) AND  (x3 = TRUE) AND  (x4 = FALSE) AND  (x5 = TRUE)) THEN 
        cstate98 := 2131; y0 := FALSE; y1 := FALSE; y2 := FALSE;  
    ELSIF ((x0 = FALSE) AND  (x1 = FALSE) AND  (x2 = FALSE) AND  (x3 = TRUE) AND  (x4 = TRUE) AND  (x5 = FALSE)) THEN 
        cstate98 := 3624; y0 := FALSE; y1 := TRUE; y2 := FALSE;  
    ELSIF ((x0 = FALSE) AND  (x1 = FALSE) AND  (x2 = FALSE) AND  (x3 = TRUE) AND  (x4 = TRUE) AND  (x5 = TRUE)) THEN 
        cstate98 := 2090; y0 := FALSE; y1 := FALSE; y2 := FALSE;  
    ELSIF ((x0 = FALSE) AND  (x1 = FALSE) AND  (x2 = TRUE) AND  (x3 = FALSE) AND  ( TRUE ) AND  (x5 = FALSE)) THEN 
        cstate98 := 2608; y0 := FALSE; y1 := TRUE; y2 := FALSE;  
    ELSIF ((x0 = FALSE) AND  (x1 = FALSE) AND  (x2 = TRUE) AND  (x3 = FALSE) AND  ( TRUE ) AND  (x5 = TRUE)) THEN 
        cstate98 := 1618; y0 := FALSE; y1 := FALSE; y2 := FALSE;  
    ELSIF ((x0 = FALSE) AND  (x1 = FALSE) AND  (x2 = TRUE) AND  (x3 = TRUE) AND  ( TRUE ) AND  ( TRUE )) OR ((x0 = FALSE) AND  (x1 = TRUE) AND  (x2 = FALSE) AND  (x3 = TRUE) AND  ( TRUE ) AND  ( TRUE )) OR ((x0 = FALSE) AND  (x1 = TRUE) AND  (x2 = TRUE) AND  ( TRUE ) AND  ( TRUE ) AND  ( TRUE )) OR ((x0 = TRUE) AND  ( TRUE ) AND  (x2 = FALSE) AND  (x3 = TRUE) AND  ( TRUE ) AND  ( TRUE )) OR ((x0 = TRUE) AND  ( TRUE ) AND  (x2 = TRUE) AND  ( TRUE ) AND  ( TRUE ) AND  ( TRUE )) THEN 
        cstate98 := 617; y0 := FALSE; y1 := FALSE; y2 := FALSE;  
    ELSIF ((x0 = FALSE) AND  (x1 = TRUE) AND  (x2 = FALSE) AND  (x3 = FALSE) AND  ( TRUE ) AND  (x5 = FALSE)) OR ((x0 = TRUE) AND  ( TRUE ) AND  (x2 = FALSE) AND  (x3 = FALSE) AND  ( TRUE ) AND  (x5 = FALSE)) THEN 
        cstate98 := 3728; y0 := FALSE; y1 := TRUE; y2 := FALSE;  
    ELSIF ((x0 = FALSE) AND  (x1 = TRUE) AND  (x2 = FALSE) AND  (x3 = FALSE) AND  ( TRUE ) AND  (x5 = TRUE)) OR ((x0 = TRUE) AND  ( TRUE ) AND  (x2 = FALSE) AND  (x3 = FALSE) AND  ( TRUE ) AND  (x5 = TRUE)) THEN 
        cstate98 := 1202; y0 := FALSE; y1 := FALSE; y2 := FALSE;  
    END_IF;
1188:
    IF ((x0 = FALSE) AND  (x1 = FALSE) AND  (x2 = FALSE) AND  (x3 = FALSE) AND  ( TRUE ) AND  (x5 = FALSE)) OR ((x0 = FALSE) AND  (x1 = FALSE) AND  (x2 = FALSE) AND  (x3 = TRUE) AND  (x4 = FALSE) AND  (x5 = FALSE)) THEN 
        cstate98 := 2212; y0 := FALSE; y1 := FALSE; y2 := FALSE;  
    ELSIF ((x0 = FALSE) AND  (x1 = FALSE) AND  (x2 = FALSE) AND  (x3 = FALSE) AND  ( TRUE ) AND  (x5 = TRUE)) OR ((x0 = FALSE) AND  (x1 = FALSE) AND  (x2 = FALSE) AND  (x3 = TRUE) AND  (x4 = FALSE) AND  (x5 = TRUE)) THEN 
        cstate98 := 2215; y0 := FALSE; y1 := FALSE; y2 := FALSE;  
    ELSIF ((x0 = FALSE) AND  (x1 = FALSE) AND  (x2 = FALSE) AND  (x3 = TRUE) AND  (x4 = TRUE) AND  (x5 = FALSE)) THEN 
        cstate98 := 236; y0 := FALSE; y1 := FALSE; y2 := TRUE;  
    ELSIF ((x0 = FALSE) AND  (x1 = FALSE) AND  (x2 = FALSE) AND  (x3 = TRUE) AND  (x4 = TRUE) AND  (x5 = TRUE)) THEN 
        cstate98 := 2190; y0 := FALSE; y1 := FALSE; y2 := FALSE;  
    ELSIF ((x0 = FALSE) AND  (x1 = FALSE) AND  (x2 = TRUE) AND  (x3 = FALSE) AND  ( TRUE ) AND  (x5 = FALSE)) THEN 
        cstate98 := 2704; y0 := FALSE; y1 := TRUE; y2 := FALSE;  
    ELSIF ((x0 = FALSE) AND  (x1 = FALSE) AND  (x2 = TRUE) AND  (x3 = FALSE) AND  ( TRUE ) AND  (x5 = TRUE)) THEN 
        cstate98 := 1714; y0 := FALSE; y1 := FALSE; y2 := FALSE;  
    ELSIF ((x0 = FALSE) AND  (x1 = FALSE) AND  (x2 = TRUE) AND  (x3 = TRUE) AND  ( TRUE ) AND  ( TRUE )) OR ((x0 = FALSE) AND  (x1 = TRUE) AND  (x2 = FALSE) AND  (x3 = TRUE) AND  ( TRUE ) AND  ( TRUE )) OR ((x0 = FALSE) AND  (x1 = TRUE) AND  (x2 = TRUE) AND  ( TRUE ) AND  ( TRUE ) AND  ( TRUE )) OR ((x0 = TRUE) AND  ( TRUE ) AND  (x2 = FALSE) AND  (x3 = TRUE) AND  ( TRUE ) AND  ( TRUE )) OR ((x0 = TRUE) AND  ( TRUE ) AND  (x2 = TRUE) AND  ( TRUE ) AND  ( TRUE ) AND  ( TRUE )) THEN 
        cstate98 := 617; y0 := FALSE; y1 := FALSE; y2 := FALSE;  
    ELSIF ((x0 = FALSE) AND  (x1 = TRUE) AND  (x2 = FALSE) AND  (x3 = FALSE) AND  ( TRUE ) AND  (x5 = FALSE)) OR ((x0 = TRUE) AND  ( TRUE ) AND  (x2 = FALSE) AND  (x3 = FALSE) AND  ( TRUE ) AND  (x5 = FALSE)) THEN 
        cstate98 := 1188; y0 := FALSE; y1 := FALSE; y2 := FALSE;  
    ELSIF ((x0 = FALSE) AND  (x1 = TRUE) AND  (x2 = FALSE) AND  (x3 = FALSE) AND  ( TRUE ) AND  (x5 = TRUE)) OR ((x0 = TRUE) AND  ( TRUE ) AND  (x2 = FALSE) AND  (x3 = FALSE) AND  ( TRUE ) AND  (x5 = TRUE)) THEN 
        cstate98 := 1190; y0 := FALSE; y1 := FALSE; y2 := FALSE;  
    END_IF;
3634:
    IF ((x0 = FALSE) AND  (x1 = FALSE) AND  (x2 = FALSE) AND  (x3 = FALSE) AND  ( TRUE ) AND  (x5 = FALSE)) OR ((x0 = FALSE) AND  (x1 = FALSE) AND  (x2 = FALSE) AND  (x3 = TRUE) AND  (x4 = FALSE) AND  (x5 = FALSE)) THEN 
        cstate98 := 3634; y0 := FALSE; y1 := TRUE; y2 := FALSE;  
    ELSIF ((x0 = FALSE) AND  (x1 = FALSE) AND  (x2 = FALSE) AND  (x3 = FALSE) AND  ( TRUE ) AND  (x5 = TRUE)) OR ((x0 = FALSE) AND  (x1 = FALSE) AND  (x2 = FALSE) AND  (x3 = TRUE) AND  (x4 = FALSE) AND  (x5 = TRUE)) THEN 
        cstate98 := 2131; y0 := FALSE; y1 := FALSE; y2 := FALSE;  
    ELSIF ((x0 = FALSE) AND  (x1 = FALSE) AND  (x2 = FALSE) AND  (x3 = TRUE) AND  (x4 = TRUE) AND  (x5 = FALSE)) THEN 
        cstate98 := 3626; y0 := FALSE; y1 := TRUE; y2 := FALSE;  
    ELSIF ((x0 = FALSE) AND  (x1 = FALSE) AND  (x2 = FALSE) AND  (x3 = TRUE) AND  (x4 = TRUE) AND  (x5 = TRUE)) THEN 
        cstate98 := 2090; y0 := FALSE; y1 := FALSE; y2 := FALSE;  
    ELSIF ((x0 = FALSE) AND  (x1 = FALSE) AND  (x2 = TRUE) AND  (x3 = FALSE) AND  ( TRUE ) AND  (x5 = FALSE)) THEN 
        cstate98 := 2610; y0 := FALSE; y1 := TRUE; y2 := FALSE;  
    ELSIF ((x0 = FALSE) AND  (x1 = FALSE) AND  (x2 = TRUE) AND  (x3 = FALSE) AND  ( TRUE ) AND  (x5 = TRUE)) THEN 
        cstate98 := 1618; y0 := FALSE; y1 := FALSE; y2 := FALSE;  
    ELSIF ((x0 = FALSE) AND  (x1 = FALSE) AND  (x2 = TRUE) AND  (x3 = TRUE) AND  ( TRUE ) AND  ( TRUE )) OR ((x0 = FALSE) AND  (x1 = TRUE) AND  (x2 = FALSE) AND  (x3 = TRUE) AND  ( TRUE ) AND  ( TRUE )) OR ((x0 = FALSE) AND  (x1 = TRUE) AND  (x2 = TRUE) AND  ( TRUE ) AND  ( TRUE ) AND  ( TRUE )) OR ((x0 = TRUE) AND  ( TRUE ) AND  (x2 = FALSE) AND  (x3 = TRUE) AND  ( TRUE ) AND  ( TRUE )) OR ((x0 = TRUE) AND  ( TRUE ) AND  (x2 = TRUE) AND  ( TRUE ) AND  ( TRUE ) AND  ( TRUE )) THEN 
        cstate98 := 617; y0 := FALSE; y1 := FALSE; y2 := FALSE;  
    ELSIF ((x0 = FALSE) AND  (x1 = TRUE) AND  (x2 = FALSE) AND  (x3 = FALSE) AND  ( TRUE ) AND  (x5 = FALSE)) OR ((x0 = TRUE) AND  ( TRUE ) AND  (x2 = FALSE) AND  (x3 = FALSE) AND  ( TRUE ) AND  (x5 = FALSE)) THEN 
        cstate98 := 3730; y0 := FALSE; y1 := TRUE; y2 := FALSE;  
    ELSIF ((x0 = FALSE) AND  (x1 = TRUE) AND  (x2 = FALSE) AND  (x3 = FALSE) AND  ( TRUE ) AND  (x5 = TRUE)) OR ((x0 = TRUE) AND  ( TRUE ) AND  (x2 = FALSE) AND  (x3 = FALSE) AND  ( TRUE ) AND  (x5 = TRUE)) THEN 
        cstate98 := 1202; y0 := FALSE; y1 := FALSE; y2 := FALSE;  
    END_IF;
2190:
    IF ((x0 = FALSE) AND  (x1 = FALSE) AND  (x2 = FALSE) AND  (x3 = FALSE) AND  ( TRUE ) AND  (x5 = FALSE)) OR ((x0 = FALSE) AND  (x1 = FALSE) AND  (x2 = FALSE) AND  (x3 = TRUE) AND  (x4 = FALSE) AND  (x5 = FALSE)) THEN 
        cstate98 := 2222; y0 := FALSE; y1 := FALSE; y2 := FALSE;  
    ELSIF ((x0 = FALSE) AND  (x1 = FALSE) AND  (x2 = FALSE) AND  (x3 = FALSE) AND  ( TRUE ) AND  (x5 = TRUE)) OR ((x0 = FALSE) AND  (x1 = FALSE) AND  (x2 = FALSE) AND  (x3 = TRUE) AND  (x4 = FALSE) AND  (x5 = TRUE)) THEN 
        cstate98 := 2223; y0 := FALSE; y1 := FALSE; y2 := FALSE;  
    ELSIF ((x0 = FALSE) AND  (x1 = FALSE) AND  (x2 = FALSE) AND  (x3 = TRUE) AND  (x4 = TRUE) AND  ( TRUE )) THEN 
        cstate98 := 2190; y0 := FALSE; y1 := FALSE; y2 := FALSE;  
    ELSIF ((x0 = FALSE) AND  (x1 = FALSE) AND  (x2 = TRUE) AND  (x3 = FALSE) AND  ( TRUE ) AND  (x5 = FALSE)) THEN 
        cstate98 := 2698; y0 := FALSE; y1 := TRUE; y2 := FALSE;  
    ELSIF ((x0 = FALSE) AND  (x1 = FALSE) AND  (x2 = TRUE) AND  (x3 = FALSE) AND  ( TRUE ) AND  (x5 = TRUE)) THEN 
        cstate98 := 1706; y0 := FALSE; y1 := FALSE; y2 := FALSE;  
    ELSIF ((x0 = FALSE) AND  (x1 = FALSE) AND  (x2 = TRUE) AND  (x3 = TRUE) AND  ( TRUE ) AND  ( TRUE )) OR ((x0 = FALSE) AND  (x1 = TRUE) AND  (x2 = FALSE) AND  (x3 = TRUE) AND  ( TRUE ) AND  ( TRUE )) OR ((x0 = FALSE) AND  (x1 = TRUE) AND  (x2 = TRUE) AND  ( TRUE ) AND  ( TRUE ) AND  ( TRUE )) OR ((x0 = TRUE) AND  ( TRUE ) AND  (x2 = FALSE) AND  (x3 = TRUE) AND  ( TRUE ) AND  ( TRUE )) OR ((x0 = TRUE) AND  ( TRUE ) AND  (x2 = TRUE) AND  ( TRUE ) AND  ( TRUE ) AND  ( TRUE )) THEN 
        cstate98 := 617; y0 := FALSE; y1 := FALSE; y2 := FALSE;  
    ELSIF ((x0 = FALSE) AND  (x1 = TRUE) AND  (x2 = FALSE) AND  (x3 = FALSE) AND  ( TRUE ) AND  (x5 = FALSE)) OR ((x0 = TRUE) AND  ( TRUE ) AND  (x2 = FALSE) AND  (x3 = FALSE) AND  ( TRUE ) AND  (x5 = FALSE)) THEN 
        cstate98 := 3214; y0 := TRUE; y1 := FALSE; y2 := FALSE;  
    ELSIF ((x0 = FALSE) AND  (x1 = TRUE) AND  (x2 = FALSE) AND  (x3 = FALSE) AND  ( TRUE ) AND  (x5 = TRUE)) OR ((x0 = TRUE) AND  ( TRUE ) AND  (x2 = FALSE) AND  (x3 = FALSE) AND  ( TRUE ) AND  (x5 = TRUE)) THEN 
        cstate98 := 1198; y0 := FALSE; y1 := FALSE; y2 := FALSE;  
    END_IF;
202:
    IF ((x0 = FALSE) AND  (x1 = FALSE) AND  (x2 = FALSE) AND  (x3 = FALSE) AND  ( TRUE ) AND  (x5 = FALSE)) OR ((x0 = FALSE) AND  (x1 = FALSE) AND  (x2 = FALSE) AND  (x3 = TRUE) AND  (x4 = FALSE) AND  (x5 = FALSE)) OR ((x0 = FALSE) AND  (x1 = FALSE) AND  (x2 = TRUE) AND  (x3 = FALSE) AND  ( TRUE ) AND  (x5 = FALSE)) THEN 
        cstate98 := 266; y0 := FALSE; y1 := FALSE; y2 := TRUE;  
    ELSIF ((x0 = FALSE) AND  (x1 = FALSE) AND  (x2 = FALSE) AND  (x3 = FALSE) AND  ( TRUE ) AND  (x5 = TRUE)) OR ((x0 = FALSE) AND  (x1 = FALSE) AND  (x2 = FALSE) AND  (x3 = TRUE) AND  (x4 = FALSE) AND  (x5 = TRUE)) THEN 
        cstate98 := 2123; y0 := FALSE; y1 := FALSE; y2 := FALSE;  
    ELSIF ((x0 = FALSE) AND  (x1 = FALSE) AND  (x2 = FALSE) AND  (x3 = TRUE) AND  (x4 = TRUE) AND  (x5 = FALSE)) THEN 
        cstate98 := 202; y0 := FALSE; y1 := FALSE; y2 := TRUE;  
    ELSIF ((x0 = FALSE) AND  (x1 = FALSE) AND  (x2 = FALSE) AND  (x3 = TRUE) AND  (x4 = TRUE) AND  (x5 = TRUE)) THEN 
        cstate98 := 2090; y0 := FALSE; y1 := FALSE; y2 := FALSE;  
    ELSIF ((x0 = FALSE) AND  (x1 = FALSE) AND  (x2 = TRUE) AND  (x3 = FALSE) AND  ( TRUE ) AND  (x5 = TRUE)) THEN 
        cstate98 := 1610; y0 := FALSE; y1 := FALSE; y2 := FALSE;  
    ELSIF ((x0 = FALSE) AND  (x1 = FALSE) AND  (x2 = TRUE) AND  (x3 = TRUE) AND  ( TRUE ) AND  ( TRUE )) OR ((x0 = FALSE) AND  (x1 = TRUE) AND  (x2 = FALSE) AND  (x3 = TRUE) AND  ( TRUE ) AND  ( TRUE )) OR ((x0 = FALSE) AND  (x1 = TRUE) AND  (x2 = TRUE) AND  ( TRUE ) AND  ( TRUE ) AND  ( TRUE )) OR ((x0 = TRUE) AND  ( TRUE ) AND  (x2 = FALSE) AND  (x3 = TRUE) AND  ( TRUE ) AND  ( TRUE )) OR ((x0 = TRUE) AND  ( TRUE ) AND  (x2 = TRUE) AND  ( TRUE ) AND  ( TRUE ) AND  ( TRUE )) THEN 
        cstate98 := 617; y0 := FALSE; y1 := FALSE; y2 := FALSE;  
    ELSIF ((x0 = FALSE) AND  (x1 = TRUE) AND  (x2 = FALSE) AND  (x3 = FALSE) AND  ( TRUE ) AND  (x5 = FALSE)) OR ((x0 = TRUE) AND  ( TRUE ) AND  (x2 = FALSE) AND  (x3 = FALSE) AND  ( TRUE ) AND  (x5 = FALSE)) THEN 
        cstate98 := 298; y0 := FALSE; y1 := FALSE; y2 := TRUE;  
    ELSIF ((x0 = FALSE) AND  (x1 = TRUE) AND  (x2 = FALSE) AND  (x3 = FALSE) AND  ( TRUE ) AND  (x5 = TRUE)) OR ((x0 = TRUE) AND  ( TRUE ) AND  (x2 = FALSE) AND  (x3 = FALSE) AND  ( TRUE ) AND  (x5 = TRUE)) THEN 
        cstate98 := 1194; y0 := FALSE; y1 := FALSE; y2 := FALSE;  
    END_IF;
300:
    IF ((x0 = FALSE) AND  (x1 = FALSE) AND  (x2 = FALSE) AND  (x3 = FALSE) AND  ( TRUE ) AND  (x5 = FALSE)) OR ((x0 = FALSE) AND  (x1 = FALSE) AND  (x2 = FALSE) AND  (x3 = TRUE) AND  (x4 = FALSE) AND  (x5 = FALSE)) OR ((x0 = FALSE) AND  (x1 = TRUE) AND  (x2 = FALSE) AND  (x3 = FALSE) AND  ( TRUE ) AND  (x5 = FALSE)) OR ((x0 = TRUE) AND  ( TRUE ) AND  (x2 = FALSE) AND  (x3 = FALSE) AND  ( TRUE ) AND  (x5 = FALSE)) THEN 
        cstate98 := 300; y0 := FALSE; y1 := FALSE; y2 := TRUE;  
    ELSIF ((x0 = FALSE) AND  (x1 = FALSE) AND  (x2 = FALSE) AND  (x3 = FALSE) AND  ( TRUE ) AND  (x5 = TRUE)) OR ((x0 = FALSE) AND  (x1 = FALSE) AND  (x2 = FALSE) AND  (x3 = TRUE) AND  (x4 = FALSE) AND  (x5 = TRUE)) THEN 
        cstate98 := 2223; y0 := FALSE; y1 := FALSE; y2 := FALSE;  
    ELSIF ((x0 = FALSE) AND  (x1 = FALSE) AND  (x2 = FALSE) AND  (x3 = TRUE) AND  (x4 = TRUE) AND  (x5 = FALSE)) THEN 
        cstate98 := 236; y0 := FALSE; y1 := FALSE; y2 := TRUE;  
    ELSIF ((x0 = FALSE) AND  (x1 = FALSE) AND  (x2 = FALSE) AND  (x3 = TRUE) AND  (x4 = TRUE) AND  (x5 = TRUE)) THEN 
        cstate98 := 2190; y0 := FALSE; y1 := FALSE; y2 := FALSE;  
    ELSIF ((x0 = FALSE) AND  (x1 = FALSE) AND  (x2 = TRUE) AND  (x3 = FALSE) AND  ( TRUE ) AND  (x5 = FALSE)) THEN 
        cstate98 := 296; y0 := FALSE; y1 := FALSE; y2 := TRUE;  
    ELSIF ((x0 = FALSE) AND  (x1 = FALSE) AND  (x2 = TRUE) AND  (x3 = FALSE) AND  ( TRUE ) AND  (x5 = TRUE)) THEN 
        cstate98 := 1706; y0 := FALSE; y1 := FALSE; y2 := FALSE;  
    ELSIF ((x0 = FALSE) AND  (x1 = FALSE) AND  (x2 = TRUE) AND  (x3 = TRUE) AND  ( TRUE ) AND  ( TRUE )) OR ((x0 = FALSE) AND  (x1 = TRUE) AND  (x2 = FALSE) AND  (x3 = TRUE) AND  ( TRUE ) AND  ( TRUE )) OR ((x0 = FALSE) AND  (x1 = TRUE) AND  (x2 = TRUE) AND  ( TRUE ) AND  ( TRUE ) AND  ( TRUE )) OR ((x0 = TRUE) AND  ( TRUE ) AND  (x2 = FALSE) AND  (x3 = TRUE) AND  ( TRUE ) AND  ( TRUE )) OR ((x0 = TRUE) AND  ( TRUE ) AND  (x2 = TRUE) AND  ( TRUE ) AND  ( TRUE ) AND  ( TRUE )) THEN 
        cstate98 := 617; y0 := FALSE; y1 := FALSE; y2 := FALSE;  
    ELSIF ((x0 = FALSE) AND  (x1 = TRUE) AND  (x2 = FALSE) AND  (x3 = FALSE) AND  ( TRUE ) AND  (x5 = TRUE)) OR ((x0 = TRUE) AND  ( TRUE ) AND  (x2 = FALSE) AND  (x3 = FALSE) AND  ( TRUE ) AND  (x5 = TRUE)) THEN 
        cstate98 := 1198; y0 := FALSE; y1 := FALSE; y2 := FALSE;  
    END_IF;
204:
    IF ((x0 = FALSE) AND  (x1 = FALSE) AND  (x2 = FALSE) AND  (x3 = FALSE) AND  ( TRUE ) AND  (x5 = FALSE)) OR ((x0 = FALSE) AND  (x1 = FALSE) AND  (x2 = FALSE) AND  (x3 = TRUE) AND  (x4 = FALSE) AND  (x5 = FALSE)) THEN 
        cstate98 := 268; y0 := FALSE; y1 := FALSE; y2 := TRUE;  
    ELSIF ((x0 = FALSE) AND  (x1 = FALSE) AND  (x2 = FALSE) AND  (x3 = FALSE) AND  ( TRUE ) AND  (x5 = TRUE)) OR ((x0 = FALSE) AND  (x1 = FALSE) AND  (x2 = FALSE) AND  (x3 = TRUE) AND  (x4 = FALSE) AND  (x5 = TRUE)) THEN 
        cstate98 := 2127; y0 := FALSE; y1 := FALSE; y2 := FALSE;  
    ELSIF ((x0 = FALSE) AND  (x1 = FALSE) AND  (x2 = FALSE) AND  (x3 = TRUE) AND  (x4 = TRUE) AND  (x5 = FALSE)) THEN 
        cstate98 := 204; y0 := FALSE; y1 := FALSE; y2 := TRUE;  
    ELSIF ((x0 = FALSE) AND  (x1 = FALSE) AND  (x2 = FALSE) AND  (x3 = TRUE) AND  (x4 = TRUE) AND  (x5 = TRUE)) THEN 
        cstate98 := 2094; y0 := FALSE; y1 := FALSE; y2 := FALSE;  
    ELSIF ((x0 = FALSE) AND  (x1 = FALSE) AND  (x2 = TRUE) AND  (x3 = FALSE) AND  ( TRUE ) AND  (x5 = FALSE)) THEN 
        cstate98 := 264; y0 := FALSE; y1 := FALSE; y2 := TRUE;  
    ELSIF ((x0 = FALSE) AND  (x1 = FALSE) AND  (x2 = TRUE) AND  (x3 = FALSE) AND  ( TRUE ) AND  (x5 = TRUE)) THEN 
        cstate98 := 1610; y0 := FALSE; y1 := FALSE; y2 := FALSE;  
    ELSIF ((x0 = FALSE) AND  (x1 = FALSE) AND  (x2 = TRUE) AND  (x3 = TRUE) AND  ( TRUE ) AND  ( TRUE )) OR ((x0 = FALSE) AND  (x1 = TRUE) AND  (x2 = FALSE) AND  (x3 = TRUE) AND  ( TRUE ) AND  ( TRUE )) OR ((x0 = FALSE) AND  (x1 = TRUE) AND  (x2 = TRUE) AND  ( TRUE ) AND  ( TRUE ) AND  ( TRUE )) OR ((x0 = TRUE) AND  ( TRUE ) AND  (x2 = FALSE) AND  (x3 = TRUE) AND  ( TRUE ) AND  ( TRUE )) OR ((x0 = TRUE) AND  ( TRUE ) AND  (x2 = TRUE) AND  ( TRUE ) AND  ( TRUE ) AND  ( TRUE )) THEN 
        cstate98 := 617; y0 := FALSE; y1 := FALSE; y2 := FALSE;  
    ELSIF ((x0 = FALSE) AND  (x1 = TRUE) AND  (x2 = FALSE) AND  (x3 = FALSE) AND  ( TRUE ) AND  (x5 = FALSE)) OR ((x0 = TRUE) AND  ( TRUE ) AND  (x2 = FALSE) AND  (x3 = FALSE) AND  ( TRUE ) AND  (x5 = FALSE)) THEN 
        cstate98 := 300; y0 := FALSE; y1 := FALSE; y2 := TRUE;  
    ELSIF ((x0 = FALSE) AND  (x1 = TRUE) AND  (x2 = FALSE) AND  (x3 = FALSE) AND  ( TRUE ) AND  (x5 = TRUE)) OR ((x0 = TRUE) AND  ( TRUE ) AND  (x2 = FALSE) AND  (x3 = FALSE) AND  ( TRUE ) AND  (x5 = TRUE)) THEN 
        cstate98 := 1198; y0 := FALSE; y1 := FALSE; y2 := FALSE;  
    END_IF;
3204:
    IF ((x0 = FALSE) AND  (x1 = FALSE) AND  (x2 = FALSE) AND  (x3 = FALSE) AND  ( TRUE ) AND  (x5 = FALSE)) OR ((x0 = FALSE) AND  (x1 = FALSE) AND  (x2 = FALSE) AND  (x3 = TRUE) AND  (x4 = FALSE) AND  (x5 = FALSE)) THEN 
        cstate98 := 4228; y0 := TRUE; y1 := FALSE; y2 := FALSE;  
    ELSIF ((x0 = FALSE) AND  (x1 = FALSE) AND  (x2 = FALSE) AND  (x3 = FALSE) AND  ( TRUE ) AND  (x5 = TRUE)) OR ((x0 = FALSE) AND  (x1 = FALSE) AND  (x2 = FALSE) AND  (x3 = TRUE) AND  (x4 = FALSE) AND  (x5 = TRUE)) THEN 
        cstate98 := 2215; y0 := FALSE; y1 := FALSE; y2 := FALSE;  
    ELSIF ((x0 = FALSE) AND  (x1 = FALSE) AND  (x2 = FALSE) AND  (x3 = TRUE) AND  (x4 = TRUE) AND  (x5 = FALSE)) THEN 
        cstate98 := 4236; y0 := TRUE; y1 := FALSE; y2 := FALSE;  
    ELSIF ((x0 = FALSE) AND  (x1 = FALSE) AND  (x2 = FALSE) AND  (x3 = TRUE) AND  (x4 = TRUE) AND  (x5 = TRUE)) THEN 
        cstate98 := 2190; y0 := FALSE; y1 := FALSE; y2 := FALSE;  
    ELSIF ((x0 = FALSE) AND  (x1 = FALSE) AND  (x2 = TRUE) AND  (x3 = FALSE) AND  ( TRUE ) AND  (x5 = FALSE)) THEN 
        cstate98 := 4240; y0 := TRUE; y1 := FALSE; y2 := FALSE;  
    ELSIF ((x0 = FALSE) AND  (x1 = FALSE) AND  (x2 = TRUE) AND  (x3 = FALSE) AND  ( TRUE ) AND  (x5 = TRUE)) THEN 
        cstate98 := 1714; y0 := FALSE; y1 := FALSE; y2 := FALSE;  
    ELSIF ((x0 = FALSE) AND  (x1 = FALSE) AND  (x2 = TRUE) AND  (x3 = TRUE) AND  ( TRUE ) AND  ( TRUE )) OR ((x0 = FALSE) AND  (x1 = TRUE) AND  (x2 = FALSE) AND  (x3 = TRUE) AND  ( TRUE ) AND  ( TRUE )) OR ((x0 = FALSE) AND  (x1 = TRUE) AND  (x2 = TRUE) AND  ( TRUE ) AND  ( TRUE ) AND  ( TRUE )) OR ((x0 = TRUE) AND  ( TRUE ) AND  (x2 = FALSE) AND  (x3 = TRUE) AND  ( TRUE ) AND  ( TRUE )) OR ((x0 = TRUE) AND  ( TRUE ) AND  (x2 = TRUE) AND  ( TRUE ) AND  ( TRUE ) AND  ( TRUE )) THEN 
        cstate98 := 617; y0 := FALSE; y1 := FALSE; y2 := FALSE;  
    ELSIF ((x0 = FALSE) AND  (x1 = TRUE) AND  (x2 = FALSE) AND  (x3 = FALSE) AND  ( TRUE ) AND  (x5 = FALSE)) OR ((x0 = TRUE) AND  ( TRUE ) AND  (x2 = FALSE) AND  (x3 = FALSE) AND  ( TRUE ) AND  (x5 = FALSE)) THEN 
        cstate98 := 3204; y0 := TRUE; y1 := FALSE; y2 := FALSE;  
    ELSIF ((x0 = FALSE) AND  (x1 = TRUE) AND  (x2 = FALSE) AND  (x3 = FALSE) AND  ( TRUE ) AND  (x5 = TRUE)) OR ((x0 = TRUE) AND  ( TRUE ) AND  (x2 = FALSE) AND  (x3 = FALSE) AND  ( TRUE ) AND  (x5 = TRUE)) THEN 
        cstate98 := 1190; y0 := FALSE; y1 := FALSE; y2 := FALSE;  
    END_IF;
302:
    IF ((x0 = FALSE) AND  (x1 = FALSE) AND  (x2 = FALSE) AND  (x3 = FALSE) AND  ( TRUE ) AND  (x5 = FALSE)) OR ((x0 = FALSE) AND  (x1 = FALSE) AND  (x2 = FALSE) AND  (x3 = TRUE) AND  (x4 = FALSE) AND  (x5 = FALSE)) OR ((x0 = FALSE) AND  (x1 = TRUE) AND  (x2 = FALSE) AND  (x3 = FALSE) AND  ( TRUE ) AND  (x5 = FALSE)) OR ((x0 = TRUE) AND  ( TRUE ) AND  (x2 = FALSE) AND  (x3 = FALSE) AND  ( TRUE ) AND  (x5 = FALSE)) THEN 
        cstate98 := 302; y0 := FALSE; y1 := FALSE; y2 := TRUE;  
    ELSIF ((x0 = FALSE) AND  (x1 = FALSE) AND  (x2 = FALSE) AND  (x3 = FALSE) AND  ( TRUE ) AND  (x5 = TRUE)) OR ((x0 = FALSE) AND  (x1 = FALSE) AND  (x2 = FALSE) AND  (x3 = TRUE) AND  (x4 = FALSE) AND  (x5 = TRUE)) THEN 
        cstate98 := 2223; y0 := FALSE; y1 := FALSE; y2 := FALSE;  
    ELSIF ((x0 = FALSE) AND  (x1 = FALSE) AND  (x2 = FALSE) AND  (x3 = TRUE) AND  (x4 = TRUE) AND  (x5 = FALSE)) THEN 
        cstate98 := 238; y0 := FALSE; y1 := FALSE; y2 := TRUE;  
    ELSIF ((x0 = FALSE) AND  (x1 = FALSE) AND  (x2 = FALSE) AND  (x3 = TRUE) AND  (x4 = TRUE) AND  (x5 = TRUE)) THEN 
        cstate98 := 2190; y0 := FALSE; y1 := FALSE; y2 := FALSE;  
    ELSIF ((x0 = FALSE) AND  (x1 = FALSE) AND  (x2 = TRUE) AND  (x3 = FALSE) AND  ( TRUE ) AND  (x5 = FALSE)) THEN 
        cstate98 := 298; y0 := FALSE; y1 := FALSE; y2 := TRUE;  
    ELSIF ((x0 = FALSE) AND  (x1 = FALSE) AND  (x2 = TRUE) AND  (x3 = FALSE) AND  ( TRUE ) AND  (x5 = TRUE)) THEN 
        cstate98 := 1706; y0 := FALSE; y1 := FALSE; y2 := FALSE;  
    ELSIF ((x0 = FALSE) AND  (x1 = FALSE) AND  (x2 = TRUE) AND  (x3 = TRUE) AND  ( TRUE ) AND  ( TRUE )) OR ((x0 = FALSE) AND  (x1 = TRUE) AND  (x2 = FALSE) AND  (x3 = TRUE) AND  ( TRUE ) AND  ( TRUE )) OR ((x0 = FALSE) AND  (x1 = TRUE) AND  (x2 = TRUE) AND  ( TRUE ) AND  ( TRUE ) AND  ( TRUE )) OR ((x0 = TRUE) AND  ( TRUE ) AND  (x2 = FALSE) AND  (x3 = TRUE) AND  ( TRUE ) AND  ( TRUE )) OR ((x0 = TRUE) AND  ( TRUE ) AND  (x2 = TRUE) AND  ( TRUE ) AND  ( TRUE ) AND  ( TRUE )) THEN 
        cstate98 := 617; y0 := FALSE; y1 := FALSE; y2 := FALSE;  
    ELSIF ((x0 = FALSE) AND  (x1 = TRUE) AND  (x2 = FALSE) AND  (x3 = FALSE) AND  ( TRUE ) AND  (x5 = TRUE)) OR ((x0 = TRUE) AND  ( TRUE ) AND  (x2 = FALSE) AND  (x3 = FALSE) AND  ( TRUE ) AND  (x5 = TRUE)) THEN 
        cstate98 := 1198; y0 := FALSE; y1 := FALSE; y2 := FALSE;  
    END_IF;
3206:
    IF ((x0 = FALSE) AND  (x1 = FALSE) AND  (x2 = FALSE) AND  (x3 = FALSE) AND  ( TRUE ) AND  (x5 = FALSE)) OR ((x0 = FALSE) AND  (x1 = FALSE) AND  (x2 = FALSE) AND  (x3 = TRUE) AND  (x4 = FALSE) AND  (x5 = FALSE)) THEN 
        cstate98 := 4230; y0 := TRUE; y1 := FALSE; y2 := FALSE;  
    ELSIF ((x0 = FALSE) AND  (x1 = FALSE) AND  (x2 = FALSE) AND  (x3 = FALSE) AND  ( TRUE ) AND  (x5 = TRUE)) OR ((x0 = FALSE) AND  (x1 = FALSE) AND  (x2 = FALSE) AND  (x3 = TRUE) AND  (x4 = FALSE) AND  (x5 = TRUE)) THEN 
        cstate98 := 2215; y0 := FALSE; y1 := FALSE; y2 := FALSE;  
    ELSIF ((x0 = FALSE) AND  (x1 = FALSE) AND  (x2 = FALSE) AND  (x3 = TRUE) AND  (x4 = TRUE) AND  (x5 = FALSE)) THEN 
        cstate98 := 4238; y0 := TRUE; y1 := FALSE; y2 := FALSE;  
    ELSIF ((x0 = FALSE) AND  (x1 = FALSE) AND  (x2 = FALSE) AND  (x3 = TRUE) AND  (x4 = TRUE) AND  (x5 = TRUE)) THEN 
        cstate98 := 2190; y0 := FALSE; y1 := FALSE; y2 := FALSE;  
    ELSIF ((x0 = FALSE) AND  (x1 = FALSE) AND  (x2 = TRUE) AND  (x3 = FALSE) AND  ( TRUE ) AND  (x5 = FALSE)) THEN 
        cstate98 := 4242; y0 := TRUE; y1 := FALSE; y2 := FALSE;  
    ELSIF ((x0 = FALSE) AND  (x1 = FALSE) AND  (x2 = TRUE) AND  (x3 = FALSE) AND  ( TRUE ) AND  (x5 = TRUE)) THEN 
        cstate98 := 1714; y0 := FALSE; y1 := FALSE; y2 := FALSE;  
    ELSIF ((x0 = FALSE) AND  (x1 = FALSE) AND  (x2 = TRUE) AND  (x3 = TRUE) AND  ( TRUE ) AND  ( TRUE )) OR ((x0 = FALSE) AND  (x1 = TRUE) AND  (x2 = FALSE) AND  (x3 = TRUE) AND  ( TRUE ) AND  ( TRUE )) OR ((x0 = FALSE) AND  (x1 = TRUE) AND  (x2 = TRUE) AND  ( TRUE ) AND  ( TRUE ) AND  ( TRUE )) OR ((x0 = TRUE) AND  ( TRUE ) AND  (x2 = FALSE) AND  (x3 = TRUE) AND  ( TRUE ) AND  ( TRUE )) OR ((x0 = TRUE) AND  ( TRUE ) AND  (x2 = TRUE) AND  ( TRUE ) AND  ( TRUE ) AND  ( TRUE )) THEN 
        cstate98 := 617; y0 := FALSE; y1 := FALSE; y2 := FALSE;  
    ELSIF ((x0 = FALSE) AND  (x1 = TRUE) AND  (x2 = FALSE) AND  (x3 = FALSE) AND  ( TRUE ) AND  (x5 = FALSE)) OR ((x0 = TRUE) AND  ( TRUE ) AND  (x2 = FALSE) AND  (x3 = FALSE) AND  ( TRUE ) AND  (x5 = FALSE)) THEN 
        cstate98 := 3206; y0 := TRUE; y1 := FALSE; y2 := FALSE;  
    ELSIF ((x0 = FALSE) AND  (x1 = TRUE) AND  (x2 = FALSE) AND  (x3 = FALSE) AND  ( TRUE ) AND  (x5 = TRUE)) OR ((x0 = TRUE) AND  ( TRUE ) AND  (x2 = FALSE) AND  (x3 = FALSE) AND  ( TRUE ) AND  (x5 = TRUE)) THEN 
        cstate98 := 1190; y0 := FALSE; y1 := FALSE; y2 := FALSE;  
    END_IF;
2122:
    IF ((x0 = FALSE) AND  (x1 = FALSE) AND  (x2 = FALSE) AND  (x3 = FALSE) AND  ( TRUE ) AND  (x5 = FALSE)) OR ((x0 = FALSE) AND  (x1 = FALSE) AND  (x2 = FALSE) AND  (x3 = TRUE) AND  (x4 = FALSE) AND  (x5 = FALSE)) THEN 
        cstate98 := 2122; y0 := FALSE; y1 := FALSE; y2 := FALSE;  
    ELSIF ((x0 = FALSE) AND  (x1 = FALSE) AND  (x2 = FALSE) AND  (x3 = FALSE) AND  ( TRUE ) AND  (x5 = TRUE)) OR ((x0 = FALSE) AND  (x1 = FALSE) AND  (x2 = FALSE) AND  (x3 = TRUE) AND  (x4 = FALSE) AND  (x5 = TRUE)) THEN 
        cstate98 := 2123; y0 := FALSE; y1 := FALSE; y2 := FALSE;  
    ELSIF ((x0 = FALSE) AND  (x1 = FALSE) AND  (x2 = FALSE) AND  (x3 = TRUE) AND  (x4 = TRUE) AND  (x5 = FALSE)) THEN 
        cstate98 := 202; y0 := FALSE; y1 := FALSE; y2 := TRUE;  
    ELSIF ((x0 = FALSE) AND  (x1 = FALSE) AND  (x2 = FALSE) AND  (x3 = TRUE) AND  (x4 = TRUE) AND  (x5 = TRUE)) THEN 
        cstate98 := 2090; y0 := FALSE; y1 := FALSE; y2 := FALSE;  
    ELSIF ((x0 = FALSE) AND  (x1 = FALSE) AND  (x2 = TRUE) AND  (x3 = FALSE) AND  ( TRUE ) AND  (x5 = FALSE)) THEN 
        cstate98 := 2602; y0 := FALSE; y1 := TRUE; y2 := FALSE;  
    ELSIF ((x0 = FALSE) AND  (x1 = FALSE) AND  (x2 = TRUE) AND  (x3 = FALSE) AND  ( TRUE ) AND  (x5 = TRUE)) THEN 
        cstate98 := 1610; y0 := FALSE; y1 := FALSE; y2 := FALSE;  
    ELSIF ((x0 = FALSE) AND  (x1 = FALSE) AND  (x2 = TRUE) AND  (x3 = TRUE) AND  ( TRUE ) AND  ( TRUE )) OR ((x0 = FALSE) AND  (x1 = TRUE) AND  (x2 = FALSE) AND  (x3 = TRUE) AND  ( TRUE ) AND  ( TRUE )) OR ((x0 = FALSE) AND  (x1 = TRUE) AND  (x2 = TRUE) AND  ( TRUE ) AND  ( TRUE ) AND  ( TRUE )) OR ((x0 = TRUE) AND  ( TRUE ) AND  (x2 = FALSE) AND  (x3 = TRUE) AND  ( TRUE ) AND  ( TRUE )) OR ((x0 = TRUE) AND  ( TRUE ) AND  (x2 = TRUE) AND  ( TRUE ) AND  ( TRUE ) AND  ( TRUE )) THEN 
        cstate98 := 617; y0 := FALSE; y1 := FALSE; y2 := FALSE;  
    ELSIF ((x0 = FALSE) AND  (x1 = TRUE) AND  (x2 = FALSE) AND  (x3 = FALSE) AND  ( TRUE ) AND  (x5 = FALSE)) OR ((x0 = TRUE) AND  ( TRUE ) AND  (x2 = FALSE) AND  (x3 = FALSE) AND  ( TRUE ) AND  (x5 = FALSE)) THEN 
        cstate98 := 3210; y0 := TRUE; y1 := FALSE; y2 := FALSE;  
    ELSIF ((x0 = FALSE) AND  (x1 = TRUE) AND  (x2 = FALSE) AND  (x3 = FALSE) AND  ( TRUE ) AND  (x5 = TRUE)) OR ((x0 = TRUE) AND  ( TRUE ) AND  (x2 = FALSE) AND  (x3 = FALSE) AND  ( TRUE ) AND  (x5 = TRUE)) THEN 
        cstate98 := 1194; y0 := FALSE; y1 := FALSE; y2 := FALSE;  
    END_IF;
200:
    IF ((x0 = FALSE) AND  (x1 = FALSE) AND  (x2 = FALSE) AND  (x3 = FALSE) AND  ( TRUE ) AND  (x5 = FALSE)) OR ((x0 = FALSE) AND  (x1 = FALSE) AND  (x2 = FALSE) AND  (x3 = TRUE) AND  (x4 = FALSE) AND  (x5 = FALSE)) OR ((x0 = FALSE) AND  (x1 = FALSE) AND  (x2 = TRUE) AND  (x3 = FALSE) AND  ( TRUE ) AND  (x5 = FALSE)) THEN 
        cstate98 := 264; y0 := FALSE; y1 := FALSE; y2 := TRUE;  
    ELSIF ((x0 = FALSE) AND  (x1 = FALSE) AND  (x2 = FALSE) AND  (x3 = FALSE) AND  ( TRUE ) AND  (x5 = TRUE)) OR ((x0 = FALSE) AND  (x1 = FALSE) AND  (x2 = FALSE) AND  (x3 = TRUE) AND  (x4 = FALSE) AND  (x5 = TRUE)) THEN 
        cstate98 := 2123; y0 := FALSE; y1 := FALSE; y2 := FALSE;  
    ELSIF ((x0 = FALSE) AND  (x1 = FALSE) AND  (x2 = FALSE) AND  (x3 = TRUE) AND  (x4 = TRUE) AND  (x5 = FALSE)) THEN 
        cstate98 := 200; y0 := FALSE; y1 := FALSE; y2 := TRUE;  
    ELSIF ((x0 = FALSE) AND  (x1 = FALSE) AND  (x2 = FALSE) AND  (x3 = TRUE) AND  (x4 = TRUE) AND  (x5 = TRUE)) THEN 
        cstate98 := 2090; y0 := FALSE; y1 := FALSE; y2 := FALSE;  
    ELSIF ((x0 = FALSE) AND  (x1 = FALSE) AND  (x2 = TRUE) AND  (x3 = FALSE) AND  ( TRUE ) AND  (x5 = TRUE)) THEN 
        cstate98 := 1610; y0 := FALSE; y1 := FALSE; y2 := FALSE;  
    ELSIF ((x0 = FALSE) AND  (x1 = FALSE) AND  (x2 = TRUE) AND  (x3 = TRUE) AND  ( TRUE ) AND  ( TRUE )) OR ((x0 = FALSE) AND  (x1 = TRUE) AND  (x2 = FALSE) AND  (x3 = TRUE) AND  ( TRUE ) AND  ( TRUE )) OR ((x0 = FALSE) AND  (x1 = TRUE) AND  (x2 = TRUE) AND  ( TRUE ) AND  ( TRUE ) AND  ( TRUE )) OR ((x0 = TRUE) AND  ( TRUE ) AND  (x2 = FALSE) AND  (x3 = TRUE) AND  ( TRUE ) AND  ( TRUE )) OR ((x0 = TRUE) AND  ( TRUE ) AND  (x2 = TRUE) AND  ( TRUE ) AND  ( TRUE ) AND  ( TRUE )) THEN 
        cstate98 := 617; y0 := FALSE; y1 := FALSE; y2 := FALSE;  
    ELSIF ((x0 = FALSE) AND  (x1 = TRUE) AND  (x2 = FALSE) AND  (x3 = FALSE) AND  ( TRUE ) AND  (x5 = FALSE)) OR ((x0 = TRUE) AND  ( TRUE ) AND  (x2 = FALSE) AND  (x3 = FALSE) AND  ( TRUE ) AND  (x5 = FALSE)) THEN 
        cstate98 := 296; y0 := FALSE; y1 := FALSE; y2 := TRUE;  
    ELSIF ((x0 = FALSE) AND  (x1 = TRUE) AND  (x2 = FALSE) AND  (x3 = FALSE) AND  ( TRUE ) AND  (x5 = TRUE)) OR ((x0 = TRUE) AND  ( TRUE ) AND  (x2 = FALSE) AND  (x3 = FALSE) AND  ( TRUE ) AND  (x5 = TRUE)) THEN 
        cstate98 := 1194; y0 := FALSE; y1 := FALSE; y2 := FALSE;  
    END_IF;
3208:
    IF ((x0 = FALSE) AND  (x1 = FALSE) AND  (x2 = FALSE) AND  ( TRUE ) AND  ( TRUE ) AND  (x5 = FALSE)) OR ((x0 = FALSE) AND  (x1 = FALSE) AND  (x2 = TRUE) AND  (x3 = FALSE) AND  ( TRUE ) AND  (x5 = FALSE)) THEN 
        cstate98 := 4232; y0 := TRUE; y1 := FALSE; y2 := FALSE;  
    ELSIF ((x0 = FALSE) AND  (x1 = FALSE) AND  (x2 = FALSE) AND  (x3 = FALSE) AND  ( TRUE ) AND  (x5 = TRUE)) OR ((x0 = FALSE) AND  (x1 = FALSE) AND  (x2 = FALSE) AND  (x3 = TRUE) AND  (x4 = FALSE) AND  (x5 = TRUE)) THEN 
        cstate98 := 2219; y0 := FALSE; y1 := FALSE; y2 := FALSE;  
    ELSIF ((x0 = FALSE) AND  (x1 = FALSE) AND  (x2 = FALSE) AND  (x3 = TRUE) AND  (x4 = TRUE) AND  (x5 = TRUE)) THEN 
        cstate98 := 2186; y0 := FALSE; y1 := FALSE; y2 := FALSE;  
    ELSIF ((x0 = FALSE) AND  (x1 = FALSE) AND  (x2 = TRUE) AND  (x3 = FALSE) AND  ( TRUE ) AND  (x5 = TRUE)) THEN 
        cstate98 := 1706; y0 := FALSE; y1 := FALSE; y2 := FALSE;  
    ELSIF ((x0 = FALSE) AND  (x1 = FALSE) AND  (x2 = TRUE) AND  (x3 = TRUE) AND  ( TRUE ) AND  ( TRUE )) OR ((x0 = FALSE) AND  (x1 = TRUE) AND  (x2 = FALSE) AND  (x3 = TRUE) AND  ( TRUE ) AND  ( TRUE )) OR ((x0 = FALSE) AND  (x1 = TRUE) AND  (x2 = TRUE) AND  ( TRUE ) AND  ( TRUE ) AND  ( TRUE )) OR ((x0 = TRUE) AND  ( TRUE ) AND  (x2 = FALSE) AND  (x3 = TRUE) AND  ( TRUE ) AND  ( TRUE )) OR ((x0 = TRUE) AND  ( TRUE ) AND  (x2 = TRUE) AND  ( TRUE ) AND  ( TRUE ) AND  ( TRUE )) THEN 
        cstate98 := 617; y0 := FALSE; y1 := FALSE; y2 := FALSE;  
    ELSIF ((x0 = FALSE) AND  (x1 = TRUE) AND  (x2 = FALSE) AND  (x3 = FALSE) AND  ( TRUE ) AND  (x5 = FALSE)) OR ((x0 = TRUE) AND  ( TRUE ) AND  (x2 = FALSE) AND  (x3 = FALSE) AND  ( TRUE ) AND  (x5 = FALSE)) THEN 
        cstate98 := 3208; y0 := TRUE; y1 := FALSE; y2 := FALSE;  
    ELSIF ((x0 = FALSE) AND  (x1 = TRUE) AND  (x2 = FALSE) AND  (x3 = FALSE) AND  ( TRUE ) AND  (x5 = TRUE)) OR ((x0 = TRUE) AND  ( TRUE ) AND  (x2 = FALSE) AND  (x3 = FALSE) AND  ( TRUE ) AND  (x5 = TRUE)) THEN 
        cstate98 := 1194; y0 := FALSE; y1 := FALSE; y2 := FALSE;  
    END_IF;
270:
    IF ((x0 = FALSE) AND  (x1 = FALSE) AND  (x2 = FALSE) AND  (x3 = FALSE) AND  ( TRUE ) AND  (x5 = FALSE)) OR ((x0 = FALSE) AND  (x1 = FALSE) AND  (x2 = FALSE) AND  (x3 = TRUE) AND  (x4 = FALSE) AND  (x5 = FALSE)) THEN 
        cstate98 := 270; y0 := FALSE; y1 := FALSE; y2 := TRUE;  
    ELSIF ((x0 = FALSE) AND  (x1 = FALSE) AND  (x2 = FALSE) AND  (x3 = FALSE) AND  ( TRUE ) AND  (x5 = TRUE)) OR ((x0 = FALSE) AND  (x1 = FALSE) AND  (x2 = FALSE) AND  (x3 = TRUE) AND  (x4 = FALSE) AND  (x5 = TRUE)) THEN 
        cstate98 := 2127; y0 := FALSE; y1 := FALSE; y2 := FALSE;  
    ELSIF ((x0 = FALSE) AND  (x1 = FALSE) AND  (x2 = FALSE) AND  (x3 = TRUE) AND  (x4 = TRUE) AND  (x5 = FALSE)) THEN 
        cstate98 := 206; y0 := FALSE; y1 := FALSE; y2 := TRUE;  
    ELSIF ((x0 = FALSE) AND  (x1 = FALSE) AND  (x2 = FALSE) AND  (x3 = TRUE) AND  (x4 = TRUE) AND  (x5 = TRUE)) THEN 
        cstate98 := 2094; y0 := FALSE; y1 := FALSE; y2 := FALSE;  
    ELSIF ((x0 = FALSE) AND  (x1 = FALSE) AND  (x2 = TRUE) AND  (x3 = FALSE) AND  ( TRUE ) AND  (x5 = FALSE)) THEN 
        cstate98 := 266; y0 := FALSE; y1 := FALSE; y2 := TRUE;  
    ELSIF ((x0 = FALSE) AND  (x1 = FALSE) AND  (x2 = TRUE) AND  (x3 = FALSE) AND  ( TRUE ) AND  (x5 = TRUE)) THEN 
        cstate98 := 1610; y0 := FALSE; y1 := FALSE; y2 := FALSE;  
    ELSIF ((x0 = FALSE) AND  (x1 = FALSE) AND  (x2 = TRUE) AND  (x3 = TRUE) AND  ( TRUE ) AND  ( TRUE )) OR ((x0 = FALSE) AND  (x1 = TRUE) AND  (x2 = FALSE) AND  (x3 = TRUE) AND  ( TRUE ) AND  ( TRUE )) OR ((x0 = FALSE) AND  (x1 = TRUE) AND  (x2 = TRUE) AND  ( TRUE ) AND  ( TRUE ) AND  ( TRUE )) OR ((x0 = TRUE) AND  ( TRUE ) AND  (x2 = FALSE) AND  (x3 = TRUE) AND  ( TRUE ) AND  ( TRUE )) OR ((x0 = TRUE) AND  ( TRUE ) AND  (x2 = TRUE) AND  ( TRUE ) AND  ( TRUE ) AND  ( TRUE )) THEN 
        cstate98 := 617; y0 := FALSE; y1 := FALSE; y2 := FALSE;  
    ELSIF ((x0 = FALSE) AND  (x1 = TRUE) AND  (x2 = FALSE) AND  (x3 = FALSE) AND  ( TRUE ) AND  (x5 = FALSE)) OR ((x0 = TRUE) AND  ( TRUE ) AND  (x2 = FALSE) AND  (x3 = FALSE) AND  ( TRUE ) AND  (x5 = FALSE)) THEN 
        cstate98 := 302; y0 := FALSE; y1 := FALSE; y2 := TRUE;  
    ELSIF ((x0 = FALSE) AND  (x1 = TRUE) AND  (x2 = FALSE) AND  (x3 = FALSE) AND  ( TRUE ) AND  (x5 = TRUE)) OR ((x0 = TRUE) AND  ( TRUE ) AND  (x2 = FALSE) AND  (x3 = FALSE) AND  ( TRUE ) AND  (x5 = TRUE)) THEN 
        cstate98 := 1198; y0 := FALSE; y1 := FALSE; y2 := FALSE;  
    END_IF;
206:
    IF ((x0 = FALSE) AND  (x1 = FALSE) AND  (x2 = FALSE) AND  (x3 = FALSE) AND  ( TRUE ) AND  (x5 = FALSE)) OR ((x0 = FALSE) AND  (x1 = FALSE) AND  (x2 = FALSE) AND  (x3 = TRUE) AND  (x4 = FALSE) AND  (x5 = FALSE)) THEN 
        cstate98 := 270; y0 := FALSE; y1 := FALSE; y2 := TRUE;  
    ELSIF ((x0 = FALSE) AND  (x1 = FALSE) AND  (x2 = FALSE) AND  (x3 = FALSE) AND  ( TRUE ) AND  (x5 = TRUE)) OR ((x0 = FALSE) AND  (x1 = FALSE) AND  (x2 = FALSE) AND  (x3 = TRUE) AND  (x4 = FALSE) AND  (x5 = TRUE)) THEN 
        cstate98 := 2127; y0 := FALSE; y1 := FALSE; y2 := FALSE;  
    ELSIF ((x0 = FALSE) AND  (x1 = FALSE) AND  (x2 = FALSE) AND  (x3 = TRUE) AND  (x4 = TRUE) AND  (x5 = FALSE)) THEN 
        cstate98 := 206; y0 := FALSE; y1 := FALSE; y2 := TRUE;  
    ELSIF ((x0 = FALSE) AND  (x1 = FALSE) AND  (x2 = FALSE) AND  (x3 = TRUE) AND  (x4 = TRUE) AND  (x5 = TRUE)) THEN 
        cstate98 := 2094; y0 := FALSE; y1 := FALSE; y2 := FALSE;  
    ELSIF ((x0 = FALSE) AND  (x1 = FALSE) AND  (x2 = TRUE) AND  (x3 = FALSE) AND  ( TRUE ) AND  (x5 = FALSE)) THEN 
        cstate98 := 266; y0 := FALSE; y1 := FALSE; y2 := TRUE;  
    ELSIF ((x0 = FALSE) AND  (x1 = FALSE) AND  (x2 = TRUE) AND  (x3 = FALSE) AND  ( TRUE ) AND  (x5 = TRUE)) THEN 
        cstate98 := 1610; y0 := FALSE; y1 := FALSE; y2 := FALSE;  
    ELSIF ((x0 = FALSE) AND  (x1 = FALSE) AND  (x2 = TRUE) AND  (x3 = TRUE) AND  ( TRUE ) AND  ( TRUE )) OR ((x0 = FALSE) AND  (x1 = TRUE) AND  (x2 = FALSE) AND  (x3 = TRUE) AND  ( TRUE ) AND  ( TRUE )) OR ((x0 = FALSE) AND  (x1 = TRUE) AND  (x2 = TRUE) AND  ( TRUE ) AND  ( TRUE ) AND  ( TRUE )) OR ((x0 = TRUE) AND  ( TRUE ) AND  (x2 = FALSE) AND  (x3 = TRUE) AND  ( TRUE ) AND  ( TRUE )) OR ((x0 = TRUE) AND  ( TRUE ) AND  (x2 = TRUE) AND  ( TRUE ) AND  ( TRUE ) AND  ( TRUE )) THEN 
        cstate98 := 617; y0 := FALSE; y1 := FALSE; y2 := FALSE;  
    ELSIF ((x0 = FALSE) AND  (x1 = TRUE) AND  (x2 = FALSE) AND  (x3 = FALSE) AND  ( TRUE ) AND  (x5 = FALSE)) OR ((x0 = TRUE) AND  ( TRUE ) AND  (x2 = FALSE) AND  (x3 = FALSE) AND  ( TRUE ) AND  (x5 = FALSE)) THEN 
        cstate98 := 302; y0 := FALSE; y1 := FALSE; y2 := TRUE;  
    ELSIF ((x0 = FALSE) AND  (x1 = TRUE) AND  (x2 = FALSE) AND  (x3 = FALSE) AND  ( TRUE ) AND  (x5 = TRUE)) OR ((x0 = TRUE) AND  ( TRUE ) AND  (x2 = FALSE) AND  (x3 = FALSE) AND  ( TRUE ) AND  (x5 = TRUE)) THEN 
        cstate98 := 1198; y0 := FALSE; y1 := FALSE; y2 := FALSE;  
    END_IF;
2610:
    IF ((x0 = FALSE) AND  (x1 = FALSE) AND  (x2 = FALSE) AND  (x3 = FALSE) AND  ( TRUE ) AND  (x5 = FALSE)) OR ((x0 = FALSE) AND  (x1 = FALSE) AND  (x2 = FALSE) AND  (x3 = TRUE) AND  (x4 = FALSE) AND  (x5 = FALSE)) THEN 
        cstate98 := 3634; y0 := FALSE; y1 := TRUE; y2 := FALSE;  
    ELSIF ((x0 = FALSE) AND  (x1 = FALSE) AND  (x2 = FALSE) AND  (x3 = FALSE) AND  ( TRUE ) AND  (x5 = TRUE)) OR ((x0 = FALSE) AND  (x1 = FALSE) AND  (x2 = FALSE) AND  (x3 = TRUE) AND  (x4 = FALSE) AND  (x5 = TRUE)) THEN 
        cstate98 := 2131; y0 := FALSE; y1 := FALSE; y2 := FALSE;  
    ELSIF ((x0 = FALSE) AND  (x1 = FALSE) AND  (x2 = FALSE) AND  (x3 = TRUE) AND  (x4 = TRUE) AND  (x5 = FALSE)) THEN 
        cstate98 := 3626; y0 := FALSE; y1 := TRUE; y2 := FALSE;  
    ELSIF ((x0 = FALSE) AND  (x1 = FALSE) AND  (x2 = FALSE) AND  (x3 = TRUE) AND  (x4 = TRUE) AND  (x5 = TRUE)) THEN 
        cstate98 := 2090; y0 := FALSE; y1 := FALSE; y2 := FALSE;  
    ELSIF ((x0 = FALSE) AND  (x1 = FALSE) AND  (x2 = TRUE) AND  (x3 = FALSE) AND  ( TRUE ) AND  (x5 = FALSE)) THEN 
        cstate98 := 2610; y0 := FALSE; y1 := TRUE; y2 := FALSE;  
    ELSIF ((x0 = FALSE) AND  (x1 = FALSE) AND  (x2 = TRUE) AND  (x3 = FALSE) AND  ( TRUE ) AND  (x5 = TRUE)) THEN 
        cstate98 := 1618; y0 := FALSE; y1 := FALSE; y2 := FALSE;  
    ELSIF ((x0 = FALSE) AND  (x1 = FALSE) AND  (x2 = TRUE) AND  (x3 = TRUE) AND  ( TRUE ) AND  ( TRUE )) OR ((x0 = FALSE) AND  (x1 = TRUE) AND  (x2 = FALSE) AND  (x3 = TRUE) AND  ( TRUE ) AND  ( TRUE )) OR ((x0 = FALSE) AND  (x1 = TRUE) AND  (x2 = TRUE) AND  ( TRUE ) AND  ( TRUE ) AND  ( TRUE )) OR ((x0 = TRUE) AND  ( TRUE ) AND  (x2 = FALSE) AND  (x3 = TRUE) AND  ( TRUE ) AND  ( TRUE )) OR ((x0 = TRUE) AND  ( TRUE ) AND  (x2 = TRUE) AND  ( TRUE ) AND  ( TRUE ) AND  ( TRUE )) THEN 
        cstate98 := 617; y0 := FALSE; y1 := FALSE; y2 := FALSE;  
    ELSIF ((x0 = FALSE) AND  (x1 = TRUE) AND  (x2 = FALSE) AND  (x3 = FALSE) AND  ( TRUE ) AND  (x5 = FALSE)) OR ((x0 = TRUE) AND  ( TRUE ) AND  (x2 = FALSE) AND  (x3 = FALSE) AND  ( TRUE ) AND  (x5 = FALSE)) THEN 
        cstate98 := 3730; y0 := FALSE; y1 := TRUE; y2 := FALSE;  
    ELSIF ((x0 = FALSE) AND  (x1 = TRUE) AND  (x2 = FALSE) AND  (x3 = FALSE) AND  ( TRUE ) AND  (x5 = TRUE)) OR ((x0 = TRUE) AND  ( TRUE ) AND  (x2 = FALSE) AND  (x3 = FALSE) AND  ( TRUE ) AND  (x5 = TRUE)) THEN 
        cstate98 := 1202; y0 := FALSE; y1 := FALSE; y2 := FALSE;  
    END_IF;
1616:
    IF ((x0 = FALSE) AND  (x1 = FALSE) AND  (x2 = FALSE) AND  (x3 = FALSE) AND  ( TRUE ) AND  (x5 = FALSE)) OR ((x0 = FALSE) AND  (x1 = FALSE) AND  (x2 = FALSE) AND  (x3 = TRUE) AND  (x4 = FALSE) AND  (x5 = FALSE)) THEN 
        cstate98 := 2128; y0 := FALSE; y1 := FALSE; y2 := FALSE;  
    ELSIF ((x0 = FALSE) AND  (x1 = FALSE) AND  (x2 = FALSE) AND  (x3 = FALSE) AND  ( TRUE ) AND  (x5 = TRUE)) OR ((x0 = FALSE) AND  (x1 = FALSE) AND  (x2 = FALSE) AND  (x3 = TRUE) AND  (x4 = FALSE) AND  (x5 = TRUE)) THEN 
        cstate98 := 2131; y0 := FALSE; y1 := FALSE; y2 := FALSE;  
    ELSIF ((x0 = FALSE) AND  (x1 = FALSE) AND  (x2 = FALSE) AND  (x3 = TRUE) AND  (x4 = TRUE) AND  (x5 = FALSE)) THEN 
        cstate98 := 200; y0 := FALSE; y1 := FALSE; y2 := TRUE;  
    ELSIF ((x0 = FALSE) AND  (x1 = FALSE) AND  (x2 = FALSE) AND  (x3 = TRUE) AND  (x4 = TRUE) AND  (x5 = TRUE)) THEN 
        cstate98 := 2090; y0 := FALSE; y1 := FALSE; y2 := FALSE;  
    ELSIF ((x0 = FALSE) AND  (x1 = FALSE) AND  (x2 = TRUE) AND  (x3 = FALSE) AND  ( TRUE ) AND  (x5 = FALSE)) THEN 
        cstate98 := 1616; y0 := FALSE; y1 := FALSE; y2 := FALSE;  
    ELSIF ((x0 = FALSE) AND  (x1 = FALSE) AND  (x2 = TRUE) AND  (x3 = FALSE) AND  ( TRUE ) AND  (x5 = TRUE)) THEN 
        cstate98 := 1618; y0 := FALSE; y1 := FALSE; y2 := FALSE;  
    ELSIF ((x0 = FALSE) AND  (x1 = FALSE) AND  (x2 = TRUE) AND  (x3 = TRUE) AND  ( TRUE ) AND  ( TRUE )) OR ((x0 = FALSE) AND  (x1 = TRUE) AND  (x2 = FALSE) AND  (x3 = TRUE) AND  ( TRUE ) AND  ( TRUE )) OR ((x0 = FALSE) AND  (x1 = TRUE) AND  (x2 = TRUE) AND  ( TRUE ) AND  ( TRUE ) AND  ( TRUE )) OR ((x0 = TRUE) AND  ( TRUE ) AND  (x2 = FALSE) AND  (x3 = TRUE) AND  ( TRUE ) AND  ( TRUE )) OR ((x0 = TRUE) AND  ( TRUE ) AND  (x2 = TRUE) AND  ( TRUE ) AND  ( TRUE ) AND  ( TRUE )) THEN 
        cstate98 := 617; y0 := FALSE; y1 := FALSE; y2 := FALSE;  
    ELSIF ((x0 = FALSE) AND  (x1 = TRUE) AND  (x2 = FALSE) AND  (x3 = FALSE) AND  ( TRUE ) AND  (x5 = FALSE)) OR ((x0 = TRUE) AND  ( TRUE ) AND  (x2 = FALSE) AND  (x3 = FALSE) AND  ( TRUE ) AND  (x5 = FALSE)) THEN 
        cstate98 := 3216; y0 := TRUE; y1 := FALSE; y2 := FALSE;  
    ELSIF ((x0 = FALSE) AND  (x1 = TRUE) AND  (x2 = FALSE) AND  (x3 = FALSE) AND  ( TRUE ) AND  (x5 = TRUE)) OR ((x0 = TRUE) AND  ( TRUE ) AND  (x2 = FALSE) AND  (x3 = FALSE) AND  ( TRUE ) AND  (x5 = TRUE)) THEN 
        cstate98 := 1202; y0 := FALSE; y1 := FALSE; y2 := FALSE;  
    END_IF;
0:
    IF ((x0 = FALSE) AND  (x1 = FALSE) AND  (x2 = FALSE) AND  (x3 = FALSE) AND  ( TRUE ) AND  (x5 = FALSE)) OR ((x0 = FALSE) AND  (x1 = FALSE) AND  (x2 = FALSE) AND  (x3 = TRUE) AND  (x4 = FALSE) AND  (x5 = FALSE)) THEN 
        cstate98 := 2116; y0 := FALSE; y1 := FALSE; y2 := FALSE;  
    ELSIF ((x0 = FALSE) AND  (x1 = FALSE) AND  (x2 = FALSE) AND  (x3 = FALSE) AND  ( TRUE ) AND  (x5 = TRUE)) OR ((x0 = FALSE) AND  (x1 = FALSE) AND  (x2 = FALSE) AND  (x3 = TRUE) AND  (x4 = FALSE) AND  (x5 = TRUE)) THEN 
        cstate98 := 2119; y0 := FALSE; y1 := FALSE; y2 := FALSE;  
    ELSIF ((x0 = FALSE) AND  (x1 = FALSE) AND  (x2 = FALSE) AND  (x3 = TRUE) AND  (x4 = TRUE) AND  (x5 = FALSE)) THEN 
        cstate98 := 2092; y0 := FALSE; y1 := FALSE; y2 := FALSE;  
    ELSIF ((x0 = FALSE) AND  (x1 = FALSE) AND  (x2 = FALSE) AND  (x3 = TRUE) AND  (x4 = TRUE) AND  (x5 = TRUE)) THEN 
        cstate98 := 2094; y0 := FALSE; y1 := FALSE; y2 := FALSE;  
    ELSIF ((x0 = FALSE) AND  (x1 = FALSE) AND  (x2 = TRUE) AND  (x3 = FALSE) AND  ( TRUE ) AND  (x5 = FALSE)) THEN 
        cstate98 := 1616; y0 := FALSE; y1 := FALSE; y2 := FALSE;  
    ELSIF ((x0 = FALSE) AND  (x1 = FALSE) AND  (x2 = TRUE) AND  (x3 = FALSE) AND  ( TRUE ) AND  (x5 = TRUE)) THEN 
        cstate98 := 1618; y0 := FALSE; y1 := FALSE; y2 := FALSE;  
    ELSIF ((x0 = FALSE) AND  (x1 = FALSE) AND  (x2 = TRUE) AND  (x3 = TRUE) AND  ( TRUE ) AND  ( TRUE )) OR ((x0 = FALSE) AND  (x1 = TRUE) AND  (x2 = FALSE) AND  (x3 = TRUE) AND  ( TRUE ) AND  ( TRUE )) OR ((x0 = FALSE) AND  (x1 = TRUE) AND  (x2 = TRUE) AND  ( TRUE ) AND  ( TRUE ) AND  ( TRUE )) OR ((x0 = TRUE) AND  ( TRUE ) AND  (x2 = FALSE) AND  (x3 = TRUE) AND  ( TRUE ) AND  ( TRUE )) OR ((x0 = TRUE) AND  ( TRUE ) AND  (x2 = TRUE) AND  ( TRUE ) AND  ( TRUE ) AND  ( TRUE )) THEN 
        cstate98 := 617; y0 := FALSE; y1 := FALSE; y2 := FALSE;  
    ELSIF ((x0 = FALSE) AND  (x1 = TRUE) AND  (x2 = FALSE) AND  (x3 = FALSE) AND  ( TRUE ) AND  (x5 = FALSE)) OR ((x0 = TRUE) AND  ( TRUE ) AND  (x2 = FALSE) AND  (x3 = FALSE) AND  ( TRUE ) AND  (x5 = FALSE)) THEN 
        cstate98 := 1188; y0 := FALSE; y1 := FALSE; y2 := FALSE;  
    ELSIF ((x0 = FALSE) AND  (x1 = TRUE) AND  (x2 = FALSE) AND  (x3 = FALSE) AND  ( TRUE ) AND  (x5 = TRUE)) OR ((x0 = TRUE) AND  ( TRUE ) AND  (x2 = FALSE) AND  (x3 = FALSE) AND  ( TRUE ) AND  (x5 = TRUE)) THEN 
        cstate98 := 1190; y0 := FALSE; y1 := FALSE; y2 := FALSE;  
    END_IF;
1714:
    IF ((x0 = FALSE) AND  (x1 = FALSE) AND  (x2 = FALSE) AND  (x3 = FALSE) AND  ( TRUE ) AND  (x5 = FALSE)) OR ((x0 = FALSE) AND  (x1 = FALSE) AND  (x2 = FALSE) AND  (x3 = TRUE) AND  (x4 = FALSE) AND  (x5 = FALSE)) THEN 
        cstate98 := 2226; y0 := FALSE; y1 := FALSE; y2 := FALSE;  
    ELSIF ((x0 = FALSE) AND  (x1 = FALSE) AND  (x2 = FALSE) AND  (x3 = FALSE) AND  ( TRUE ) AND  (x5 = TRUE)) OR ((x0 = FALSE) AND  (x1 = FALSE) AND  (x2 = FALSE) AND  (x3 = TRUE) AND  (x4 = FALSE) AND  (x5 = TRUE)) THEN 
        cstate98 := 2227; y0 := FALSE; y1 := FALSE; y2 := FALSE;  
    ELSIF ((x0 = FALSE) AND  (x1 = FALSE) AND  (x2 = FALSE) AND  (x3 = TRUE) AND  (x4 = TRUE) AND  (x5 = FALSE)) THEN 
        cstate98 := 234; y0 := FALSE; y1 := FALSE; y2 := TRUE;  
    ELSIF ((x0 = FALSE) AND  (x1 = FALSE) AND  (x2 = FALSE) AND  (x3 = TRUE) AND  (x4 = TRUE) AND  (x5 = TRUE)) THEN 
        cstate98 := 2186; y0 := FALSE; y1 := FALSE; y2 := FALSE;  
    ELSIF ((x0 = FALSE) AND  (x1 = FALSE) AND  (x2 = TRUE) AND  (x3 = FALSE) AND  ( TRUE ) AND  ( TRUE )) THEN 
        cstate98 := 1714; y0 := FALSE; y1 := FALSE; y2 := FALSE;  
    ELSIF ((x0 = FALSE) AND  (x1 = FALSE) AND  (x2 = TRUE) AND  (x3 = TRUE) AND  ( TRUE ) AND  ( TRUE )) OR ((x0 = FALSE) AND  (x1 = TRUE) AND  (x2 = FALSE) AND  (x3 = TRUE) AND  ( TRUE ) AND  ( TRUE )) OR ((x0 = FALSE) AND  (x1 = TRUE) AND  (x2 = TRUE) AND  ( TRUE ) AND  ( TRUE ) AND  ( TRUE )) OR ((x0 = TRUE) AND  ( TRUE ) AND  (x2 = FALSE) AND  (x3 = TRUE) AND  ( TRUE ) AND  ( TRUE )) OR ((x0 = TRUE) AND  ( TRUE ) AND  (x2 = TRUE) AND  ( TRUE ) AND  ( TRUE ) AND  ( TRUE )) THEN 
        cstate98 := 617; y0 := FALSE; y1 := FALSE; y2 := FALSE;  
    ELSIF ((x0 = FALSE) AND  (x1 = TRUE) AND  (x2 = FALSE) AND  (x3 = FALSE) AND  ( TRUE ) AND  (x5 = FALSE)) OR ((x0 = TRUE) AND  ( TRUE ) AND  (x2 = FALSE) AND  (x3 = FALSE) AND  ( TRUE ) AND  (x5 = FALSE)) THEN 
        cstate98 := 3218; y0 := TRUE; y1 := FALSE; y2 := FALSE;  
    ELSIF ((x0 = FALSE) AND  (x1 = TRUE) AND  (x2 = FALSE) AND  (x3 = FALSE) AND  ( TRUE ) AND  (x5 = TRUE)) OR ((x0 = TRUE) AND  ( TRUE ) AND  (x2 = FALSE) AND  (x3 = FALSE) AND  ( TRUE ) AND  (x5 = TRUE)) THEN 
        cstate98 := 1202; y0 := FALSE; y1 := FALSE; y2 := FALSE;  
    END_IF;
2219:
    IF ((x0 = FALSE) AND  (x1 = FALSE) AND  (x2 = FALSE) AND  (x3 = FALSE) AND  ( TRUE ) AND  ( TRUE )) OR ((x0 = FALSE) AND  (x1 = FALSE) AND  (x2 = FALSE) AND  (x3 = TRUE) AND  (x4 = FALSE) AND  ( TRUE )) THEN 
        cstate98 := 2219; y0 := FALSE; y1 := FALSE; y2 := FALSE;  
    ELSIF ((x0 = FALSE) AND  (x1 = FALSE) AND  (x2 = FALSE) AND  (x3 = TRUE) AND  (x4 = TRUE) AND  (x5 = FALSE)) THEN 
        cstate98 := 234; y0 := FALSE; y1 := FALSE; y2 := TRUE;  
    ELSIF ((x0 = FALSE) AND  (x1 = FALSE) AND  (x2 = FALSE) AND  (x3 = TRUE) AND  (x4 = TRUE) AND  (x5 = TRUE)) THEN 
        cstate98 := 2186; y0 := FALSE; y1 := FALSE; y2 := FALSE;  
    ELSIF ((x0 = FALSE) AND  (x1 = FALSE) AND  (x2 = TRUE) AND  (x3 = FALSE) AND  ( TRUE ) AND  (x5 = FALSE)) THEN 
        cstate98 := 2698; y0 := FALSE; y1 := TRUE; y2 := FALSE;  
    ELSIF ((x0 = FALSE) AND  (x1 = FALSE) AND  (x2 = TRUE) AND  (x3 = FALSE) AND  ( TRUE ) AND  (x5 = TRUE)) THEN 
        cstate98 := 1706; y0 := FALSE; y1 := FALSE; y2 := FALSE;  
    ELSIF ((x0 = FALSE) AND  (x1 = FALSE) AND  (x2 = TRUE) AND  (x3 = TRUE) AND  ( TRUE ) AND  ( TRUE )) OR ((x0 = FALSE) AND  (x1 = TRUE) AND  (x2 = FALSE) AND  (x3 = TRUE) AND  ( TRUE ) AND  ( TRUE )) OR ((x0 = FALSE) AND  (x1 = TRUE) AND  (x2 = TRUE) AND  ( TRUE ) AND  ( TRUE ) AND  ( TRUE )) OR ((x0 = TRUE) AND  ( TRUE ) AND  (x2 = FALSE) AND  (x3 = TRUE) AND  ( TRUE ) AND  ( TRUE )) OR ((x0 = TRUE) AND  ( TRUE ) AND  (x2 = TRUE) AND  ( TRUE ) AND  ( TRUE ) AND  ( TRUE )) THEN 
        cstate98 := 617; y0 := FALSE; y1 := FALSE; y2 := FALSE;  
    ELSIF ((x0 = FALSE) AND  (x1 = TRUE) AND  (x2 = FALSE) AND  (x3 = FALSE) AND  ( TRUE ) AND  (x5 = FALSE)) OR ((x0 = TRUE) AND  ( TRUE ) AND  (x2 = FALSE) AND  (x3 = FALSE) AND  ( TRUE ) AND  (x5 = FALSE)) THEN 
        cstate98 := 3210; y0 := TRUE; y1 := FALSE; y2 := FALSE;  
    ELSIF ((x0 = FALSE) AND  (x1 = TRUE) AND  (x2 = FALSE) AND  (x3 = FALSE) AND  ( TRUE ) AND  (x5 = TRUE)) OR ((x0 = TRUE) AND  ( TRUE ) AND  (x2 = FALSE) AND  (x3 = FALSE) AND  ( TRUE ) AND  (x5 = TRUE)) THEN 
        cstate98 := 1194; y0 := FALSE; y1 := FALSE; y2 := FALSE;  
    END_IF;
1618:
    IF ((x0 = FALSE) AND  (x1 = FALSE) AND  (x2 = FALSE) AND  (x3 = FALSE) AND  ( TRUE ) AND  (x5 = FALSE)) OR ((x0 = FALSE) AND  (x1 = FALSE) AND  (x2 = FALSE) AND  (x3 = TRUE) AND  (x4 = FALSE) AND  (x5 = FALSE)) THEN 
        cstate98 := 2130; y0 := FALSE; y1 := FALSE; y2 := FALSE;  
    ELSIF ((x0 = FALSE) AND  (x1 = FALSE) AND  (x2 = FALSE) AND  (x3 = FALSE) AND  ( TRUE ) AND  (x5 = TRUE)) OR ((x0 = FALSE) AND  (x1 = FALSE) AND  (x2 = FALSE) AND  (x3 = TRUE) AND  (x4 = FALSE) AND  (x5 = TRUE)) THEN 
        cstate98 := 2131; y0 := FALSE; y1 := FALSE; y2 := FALSE;  
    ELSIF ((x0 = FALSE) AND  (x1 = FALSE) AND  (x2 = FALSE) AND  (x3 = TRUE) AND  (x4 = TRUE) AND  (x5 = FALSE)) THEN 
        cstate98 := 202; y0 := FALSE; y1 := FALSE; y2 := TRUE;  
    ELSIF ((x0 = FALSE) AND  (x1 = FALSE) AND  (x2 = FALSE) AND  (x3 = TRUE) AND  (x4 = TRUE) AND  (x5 = TRUE)) THEN 
        cstate98 := 2090; y0 := FALSE; y1 := FALSE; y2 := FALSE;  
    ELSIF ((x0 = FALSE) AND  (x1 = FALSE) AND  (x2 = TRUE) AND  (x3 = FALSE) AND  ( TRUE ) AND  ( TRUE )) THEN 
        cstate98 := 1618; y0 := FALSE; y1 := FALSE; y2 := FALSE;  
    ELSIF ((x0 = FALSE) AND  (x1 = FALSE) AND  (x2 = TRUE) AND  (x3 = TRUE) AND  ( TRUE ) AND  ( TRUE )) OR ((x0 = FALSE) AND  (x1 = TRUE) AND  (x2 = FALSE) AND  (x3 = TRUE) AND  ( TRUE ) AND  ( TRUE )) OR ((x0 = FALSE) AND  (x1 = TRUE) AND  (x2 = TRUE) AND  ( TRUE ) AND  ( TRUE ) AND  ( TRUE )) OR ((x0 = TRUE) AND  ( TRUE ) AND  (x2 = FALSE) AND  (x3 = TRUE) AND  ( TRUE ) AND  ( TRUE )) OR ((x0 = TRUE) AND  ( TRUE ) AND  (x2 = TRUE) AND  ( TRUE ) AND  ( TRUE ) AND  ( TRUE )) THEN 
        cstate98 := 617; y0 := FALSE; y1 := FALSE; y2 := FALSE;  
    ELSIF ((x0 = FALSE) AND  (x1 = TRUE) AND  (x2 = FALSE) AND  (x3 = FALSE) AND  ( TRUE ) AND  (x5 = FALSE)) OR ((x0 = TRUE) AND  ( TRUE ) AND  (x2 = FALSE) AND  (x3 = FALSE) AND  ( TRUE ) AND  (x5 = FALSE)) THEN 
        cstate98 := 3218; y0 := TRUE; y1 := FALSE; y2 := FALSE;  
    ELSIF ((x0 = FALSE) AND  (x1 = TRUE) AND  (x2 = FALSE) AND  (x3 = FALSE) AND  ( TRUE ) AND  (x5 = TRUE)) OR ((x0 = TRUE) AND  ( TRUE ) AND  (x2 = FALSE) AND  (x3 = FALSE) AND  ( TRUE ) AND  (x5 = TRUE)) THEN 
        cstate98 := 1202; y0 := FALSE; y1 := FALSE; y2 := FALSE;  
    END_IF;
232:
    IF ((x0 = FALSE) AND  (x1 = FALSE) AND  (x2 = FALSE) AND  (x3 = FALSE) AND  ( TRUE ) AND  (x5 = FALSE)) OR ((x0 = FALSE) AND  (x1 = FALSE) AND  (x2 = FALSE) AND  (x3 = TRUE) AND  (x4 = FALSE) AND  (x5 = FALSE)) OR ((x0 = FALSE) AND  (x1 = FALSE) AND  (x2 = TRUE) AND  (x3 = FALSE) AND  ( TRUE ) AND  (x5 = FALSE)) OR ((x0 = FALSE) AND  (x1 = TRUE) AND  (x2 = FALSE) AND  (x3 = FALSE) AND  ( TRUE ) AND  (x5 = FALSE)) OR ((x0 = TRUE) AND  ( TRUE ) AND  (x2 = FALSE) AND  (x3 = FALSE) AND  ( TRUE ) AND  (x5 = FALSE)) THEN 
        cstate98 := 296; y0 := FALSE; y1 := FALSE; y2 := TRUE;  
    ELSIF ((x0 = FALSE) AND  (x1 = FALSE) AND  (x2 = FALSE) AND  (x3 = FALSE) AND  ( TRUE ) AND  (x5 = TRUE)) OR ((x0 = FALSE) AND  (x1 = FALSE) AND  (x2 = FALSE) AND  (x3 = TRUE) AND  (x4 = FALSE) AND  (x5 = TRUE)) THEN 
        cstate98 := 2219; y0 := FALSE; y1 := FALSE; y2 := FALSE;  
    ELSIF ((x0 = FALSE) AND  (x1 = FALSE) AND  (x2 = FALSE) AND  (x3 = TRUE) AND  (x4 = TRUE) AND  (x5 = FALSE)) THEN 
        cstate98 := 232; y0 := FALSE; y1 := FALSE; y2 := TRUE;  
    ELSIF ((x0 = FALSE) AND  (x1 = FALSE) AND  (x2 = FALSE) AND  (x3 = TRUE) AND  (x4 = TRUE) AND  (x5 = TRUE)) THEN 
        cstate98 := 2186; y0 := FALSE; y1 := FALSE; y2 := FALSE;  
    ELSIF ((x0 = FALSE) AND  (x1 = FALSE) AND  (x2 = TRUE) AND  (x3 = FALSE) AND  ( TRUE ) AND  (x5 = TRUE)) THEN 
        cstate98 := 1706; y0 := FALSE; y1 := FALSE; y2 := FALSE;  
    ELSIF ((x0 = FALSE) AND  (x1 = FALSE) AND  (x2 = TRUE) AND  (x3 = TRUE) AND  ( TRUE ) AND  ( TRUE )) OR ((x0 = FALSE) AND  (x1 = TRUE) AND  (x2 = FALSE) AND  (x3 = TRUE) AND  ( TRUE ) AND  ( TRUE )) OR ((x0 = FALSE) AND  (x1 = TRUE) AND  (x2 = TRUE) AND  ( TRUE ) AND  ( TRUE ) AND  ( TRUE )) OR ((x0 = TRUE) AND  ( TRUE ) AND  (x2 = FALSE) AND  (x3 = TRUE) AND  ( TRUE ) AND  ( TRUE )) OR ((x0 = TRUE) AND  ( TRUE ) AND  (x2 = TRUE) AND  ( TRUE ) AND  ( TRUE ) AND  ( TRUE )) THEN 
        cstate98 := 617; y0 := FALSE; y1 := FALSE; y2 := FALSE;  
    ELSIF ((x0 = FALSE) AND  (x1 = TRUE) AND  (x2 = FALSE) AND  (x3 = FALSE) AND  ( TRUE ) AND  (x5 = TRUE)) OR ((x0 = TRUE) AND  ( TRUE ) AND  (x2 = FALSE) AND  (x3 = FALSE) AND  ( TRUE ) AND  (x5 = TRUE)) THEN 
        cstate98 := 1194; y0 := FALSE; y1 := FALSE; y2 := FALSE;  
    END_IF;
2215:
    IF ((x0 = FALSE) AND  (x1 = FALSE) AND  (x2 = FALSE) AND  (x3 = FALSE) AND  ( TRUE ) AND  ( TRUE )) OR ((x0 = FALSE) AND  (x1 = FALSE) AND  (x2 = FALSE) AND  (x3 = TRUE) AND  (x4 = FALSE) AND  ( TRUE )) THEN 
        cstate98 := 2215; y0 := FALSE; y1 := FALSE; y2 := FALSE;  
    ELSIF ((x0 = FALSE) AND  (x1 = FALSE) AND  (x2 = FALSE) AND  (x3 = TRUE) AND  (x4 = TRUE) AND  (x5 = FALSE)) THEN 
        cstate98 := 238; y0 := FALSE; y1 := FALSE; y2 := TRUE;  
    ELSIF ((x0 = FALSE) AND  (x1 = FALSE) AND  (x2 = FALSE) AND  (x3 = TRUE) AND  (x4 = TRUE) AND  (x5 = TRUE)) THEN 
        cstate98 := 2190; y0 := FALSE; y1 := FALSE; y2 := FALSE;  
    ELSIF ((x0 = FALSE) AND  (x1 = FALSE) AND  (x2 = TRUE) AND  (x3 = FALSE) AND  ( TRUE ) AND  (x5 = FALSE)) THEN 
        cstate98 := 2706; y0 := FALSE; y1 := TRUE; y2 := FALSE;  
    ELSIF ((x0 = FALSE) AND  (x1 = FALSE) AND  (x2 = TRUE) AND  (x3 = FALSE) AND  ( TRUE ) AND  (x5 = TRUE)) THEN 
        cstate98 := 1714; y0 := FALSE; y1 := FALSE; y2 := FALSE;  
    ELSIF ((x0 = FALSE) AND  (x1 = FALSE) AND  (x2 = TRUE) AND  (x3 = TRUE) AND  ( TRUE ) AND  ( TRUE )) OR ((x0 = FALSE) AND  (x1 = TRUE) AND  (x2 = FALSE) AND  (x3 = TRUE) AND  ( TRUE ) AND  ( TRUE )) OR ((x0 = FALSE) AND  (x1 = TRUE) AND  (x2 = TRUE) AND  ( TRUE ) AND  ( TRUE ) AND  ( TRUE )) OR ((x0 = TRUE) AND  ( TRUE ) AND  (x2 = FALSE) AND  (x3 = TRUE) AND  ( TRUE ) AND  ( TRUE )) OR ((x0 = TRUE) AND  ( TRUE ) AND  (x2 = TRUE) AND  ( TRUE ) AND  ( TRUE ) AND  ( TRUE )) THEN 
        cstate98 := 617; y0 := FALSE; y1 := FALSE; y2 := FALSE;  
    ELSIF ((x0 = FALSE) AND  (x1 = TRUE) AND  (x2 = FALSE) AND  (x3 = FALSE) AND  ( TRUE ) AND  (x5 = FALSE)) OR ((x0 = TRUE) AND  ( TRUE ) AND  (x2 = FALSE) AND  (x3 = FALSE) AND  ( TRUE ) AND  (x5 = FALSE)) THEN 
        cstate98 := 3206; y0 := TRUE; y1 := FALSE; y2 := FALSE;  
    ELSIF ((x0 = FALSE) AND  (x1 = TRUE) AND  (x2 = FALSE) AND  (x3 = FALSE) AND  ( TRUE ) AND  (x5 = TRUE)) OR ((x0 = TRUE) AND  ( TRUE ) AND  (x2 = FALSE) AND  (x3 = FALSE) AND  ( TRUE ) AND  (x5 = TRUE)) THEN 
        cstate98 := 1190; y0 := FALSE; y1 := FALSE; y2 := FALSE;  
    END_IF;
2218:
    IF ((x0 = FALSE) AND  (x1 = FALSE) AND  (x2 = FALSE) AND  (x3 = FALSE) AND  ( TRUE ) AND  (x5 = FALSE)) OR ((x0 = FALSE) AND  (x1 = FALSE) AND  (x2 = FALSE) AND  (x3 = TRUE) AND  (x4 = FALSE) AND  (x5 = FALSE)) THEN 
        cstate98 := 2218; y0 := FALSE; y1 := FALSE; y2 := FALSE;  
    ELSIF ((x0 = FALSE) AND  (x1 = FALSE) AND  (x2 = FALSE) AND  (x3 = FALSE) AND  ( TRUE ) AND  (x5 = TRUE)) OR ((x0 = FALSE) AND  (x1 = FALSE) AND  (x2 = FALSE) AND  (x3 = TRUE) AND  (x4 = FALSE) AND  (x5 = TRUE)) THEN 
        cstate98 := 2219; y0 := FALSE; y1 := FALSE; y2 := FALSE;  
    ELSIF ((x0 = FALSE) AND  (x1 = FALSE) AND  (x2 = FALSE) AND  (x3 = TRUE) AND  (x4 = TRUE) AND  (x5 = FALSE)) THEN 
        cstate98 := 234; y0 := FALSE; y1 := FALSE; y2 := TRUE;  
    ELSIF ((x0 = FALSE) AND  (x1 = FALSE) AND  (x2 = FALSE) AND  (x3 = TRUE) AND  (x4 = TRUE) AND  (x5 = TRUE)) THEN 
        cstate98 := 2186; y0 := FALSE; y1 := FALSE; y2 := FALSE;  
    ELSIF ((x0 = FALSE) AND  (x1 = FALSE) AND  (x2 = TRUE) AND  (x3 = FALSE) AND  ( TRUE ) AND  (x5 = FALSE)) THEN 
        cstate98 := 2698; y0 := FALSE; y1 := TRUE; y2 := FALSE;  
    ELSIF ((x0 = FALSE) AND  (x1 = FALSE) AND  (x2 = TRUE) AND  (x3 = FALSE) AND  ( TRUE ) AND  (x5 = TRUE)) THEN 
        cstate98 := 1706; y0 := FALSE; y1 := FALSE; y2 := FALSE;  
    ELSIF ((x0 = FALSE) AND  (x1 = FALSE) AND  (x2 = TRUE) AND  (x3 = TRUE) AND  ( TRUE ) AND  ( TRUE )) OR ((x0 = FALSE) AND  (x1 = TRUE) AND  (x2 = FALSE) AND  (x3 = TRUE) AND  ( TRUE ) AND  ( TRUE )) OR ((x0 = FALSE) AND  (x1 = TRUE) AND  (x2 = TRUE) AND  ( TRUE ) AND  ( TRUE ) AND  ( TRUE )) OR ((x0 = TRUE) AND  ( TRUE ) AND  (x2 = FALSE) AND  (x3 = TRUE) AND  ( TRUE ) AND  ( TRUE )) OR ((x0 = TRUE) AND  ( TRUE ) AND  (x2 = TRUE) AND  ( TRUE ) AND  ( TRUE ) AND  ( TRUE )) THEN 
        cstate98 := 617; y0 := FALSE; y1 := FALSE; y2 := FALSE;  
    ELSIF ((x0 = FALSE) AND  (x1 = TRUE) AND  (x2 = FALSE) AND  (x3 = FALSE) AND  ( TRUE ) AND  (x5 = FALSE)) OR ((x0 = TRUE) AND  ( TRUE ) AND  (x2 = FALSE) AND  (x3 = FALSE) AND  ( TRUE ) AND  (x5 = FALSE)) THEN 
        cstate98 := 3210; y0 := TRUE; y1 := FALSE; y2 := FALSE;  
    ELSIF ((x0 = FALSE) AND  (x1 = TRUE) AND  (x2 = FALSE) AND  (x3 = FALSE) AND  ( TRUE ) AND  (x5 = TRUE)) OR ((x0 = TRUE) AND  ( TRUE ) AND  (x2 = FALSE) AND  (x3 = FALSE) AND  ( TRUE ) AND  (x5 = TRUE)) THEN 
        cstate98 := 1194; y0 := FALSE; y1 := FALSE; y2 := FALSE;  
    END_IF;
234:
    IF ((x0 = FALSE) AND  (x1 = FALSE) AND  (x2 = FALSE) AND  (x3 = FALSE) AND  ( TRUE ) AND  (x5 = FALSE)) OR ((x0 = FALSE) AND  (x1 = FALSE) AND  (x2 = FALSE) AND  (x3 = TRUE) AND  (x4 = FALSE) AND  (x5 = FALSE)) OR ((x0 = FALSE) AND  (x1 = FALSE) AND  (x2 = TRUE) AND  (x3 = FALSE) AND  ( TRUE ) AND  (x5 = FALSE)) OR ((x0 = FALSE) AND  (x1 = TRUE) AND  (x2 = FALSE) AND  (x3 = FALSE) AND  ( TRUE ) AND  (x5 = FALSE)) OR ((x0 = TRUE) AND  ( TRUE ) AND  (x2 = FALSE) AND  (x3 = FALSE) AND  ( TRUE ) AND  (x5 = FALSE)) THEN 
        cstate98 := 298; y0 := FALSE; y1 := FALSE; y2 := TRUE;  
    ELSIF ((x0 = FALSE) AND  (x1 = FALSE) AND  (x2 = FALSE) AND  (x3 = FALSE) AND  ( TRUE ) AND  (x5 = TRUE)) OR ((x0 = FALSE) AND  (x1 = FALSE) AND  (x2 = FALSE) AND  (x3 = TRUE) AND  (x4 = FALSE) AND  (x5 = TRUE)) THEN 
        cstate98 := 2219; y0 := FALSE; y1 := FALSE; y2 := FALSE;  
    ELSIF ((x0 = FALSE) AND  (x1 = FALSE) AND  (x2 = FALSE) AND  (x3 = TRUE) AND  (x4 = TRUE) AND  (x5 = FALSE)) THEN 
        cstate98 := 234; y0 := FALSE; y1 := FALSE; y2 := TRUE;  
    ELSIF ((x0 = FALSE) AND  (x1 = FALSE) AND  (x2 = FALSE) AND  (x3 = TRUE) AND  (x4 = TRUE) AND  (x5 = TRUE)) THEN 
        cstate98 := 2186; y0 := FALSE; y1 := FALSE; y2 := FALSE;  
    ELSIF ((x0 = FALSE) AND  (x1 = FALSE) AND  (x2 = TRUE) AND  (x3 = FALSE) AND  ( TRUE ) AND  (x5 = TRUE)) THEN 
        cstate98 := 1706; y0 := FALSE; y1 := FALSE; y2 := FALSE;  
    ELSIF ((x0 = FALSE) AND  (x1 = FALSE) AND  (x2 = TRUE) AND  (x3 = TRUE) AND  ( TRUE ) AND  ( TRUE )) OR ((x0 = FALSE) AND  (x1 = TRUE) AND  (x2 = FALSE) AND  (x3 = TRUE) AND  ( TRUE ) AND  ( TRUE )) OR ((x0 = FALSE) AND  (x1 = TRUE) AND  (x2 = TRUE) AND  ( TRUE ) AND  ( TRUE ) AND  ( TRUE )) OR ((x0 = TRUE) AND  ( TRUE ) AND  (x2 = FALSE) AND  (x3 = TRUE) AND  ( TRUE ) AND  ( TRUE )) OR ((x0 = TRUE) AND  ( TRUE ) AND  (x2 = TRUE) AND  ( TRUE ) AND  ( TRUE ) AND  ( TRUE )) THEN 
        cstate98 := 617; y0 := FALSE; y1 := FALSE; y2 := FALSE;  
    ELSIF ((x0 = FALSE) AND  (x1 = TRUE) AND  (x2 = FALSE) AND  (x3 = FALSE) AND  ( TRUE ) AND  (x5 = TRUE)) OR ((x0 = TRUE) AND  ( TRUE ) AND  (x2 = FALSE) AND  (x3 = FALSE) AND  ( TRUE ) AND  (x5 = TRUE)) THEN 
        cstate98 := 1194; y0 := FALSE; y1 := FALSE; y2 := FALSE;  
    END_IF;
2116:
    IF ((x0 = FALSE) AND  (x1 = FALSE) AND  (x2 = FALSE) AND  (x3 = FALSE) AND  ( TRUE ) AND  (x5 = FALSE)) OR ((x0 = FALSE) AND  (x1 = FALSE) AND  (x2 = FALSE) AND  (x3 = TRUE) AND  (x4 = FALSE) AND  (x5 = FALSE)) THEN 
        cstate98 := 2116; y0 := FALSE; y1 := FALSE; y2 := FALSE;  
    ELSIF ((x0 = FALSE) AND  (x1 = FALSE) AND  (x2 = FALSE) AND  (x3 = FALSE) AND  ( TRUE ) AND  (x5 = TRUE)) OR ((x0 = FALSE) AND  (x1 = FALSE) AND  (x2 = FALSE) AND  (x3 = TRUE) AND  (x4 = FALSE) AND  (x5 = TRUE)) THEN 
        cstate98 := 2119; y0 := FALSE; y1 := FALSE; y2 := FALSE;  
    ELSIF ((x0 = FALSE) AND  (x1 = FALSE) AND  (x2 = FALSE) AND  (x3 = TRUE) AND  (x4 = TRUE) AND  (x5 = FALSE)) THEN 
        cstate98 := 204; y0 := FALSE; y1 := FALSE; y2 := TRUE;  
    ELSIF ((x0 = FALSE) AND  (x1 = FALSE) AND  (x2 = FALSE) AND  (x3 = TRUE) AND  (x4 = TRUE) AND  (x5 = TRUE)) THEN 
        cstate98 := 2094; y0 := FALSE; y1 := FALSE; y2 := FALSE;  
    ELSIF ((x0 = FALSE) AND  (x1 = FALSE) AND  (x2 = TRUE) AND  (x3 = FALSE) AND  ( TRUE ) AND  (x5 = FALSE)) THEN 
        cstate98 := 2608; y0 := FALSE; y1 := TRUE; y2 := FALSE;  
    ELSIF ((x0 = FALSE) AND  (x1 = FALSE) AND  (x2 = TRUE) AND  (x3 = FALSE) AND  ( TRUE ) AND  (x5 = TRUE)) THEN 
        cstate98 := 1618; y0 := FALSE; y1 := FALSE; y2 := FALSE;  
